   #FRK_CfgSetWalk_DeclarationUnit := FALSE;
   IF #Phase = 1 THEN
       #ConfigStageParCfg := #ParCfg;
   END_IF;
   IF #Phase = 1 THEN
       #ConfigStageStationCfg := #StationCfg;
   END_IF;
   IF "FRK_SetRuntime".Work[#RootIndex].Payload.Info.Kind = 0 THEN
       "FRK_CfgDef_DeclarationUnit"(FieldIndex := 1);
       "FRK_SetRuntime".Work[#RootIndex].RejectScope := #Status.Name;
       "FRK_SetRuntime".Work[#RootIndex].RejectKey := "FRK_ConfigScratch".Entry.WriteKey;
       IF #Phase = 0 THEN
           IF #Access.CurrentLevel < MAX(IN1 := #Access.Policy.Required[0], IN2 := "FRK_ConfigScratch".MinRead) THEN
               RETURN;
           END_IF;
           #Ok := "FRK_ConfigGet"(Scope := #Status.Name, ModelCode := "FRK_SetRuntime".Work[#RootIndex].Payload.Info.ModelCode);
           IF NOT #Ok OR "FRK_SetRuntime".Work[#RootIndex].Payload.Info.RecordCount >= 24 THEN
               RETURN;
           END_IF;
           #Slot := "FRK_SetRuntime".Work[#RootIndex].Payload.Info.RecordCount + 1;
           "FRK_SetRuntime".Work[#RootIndex].Payload.Records[#Slot].Scope := #Status.Name;
           "FRK_SetRuntime".Work[#RootIndex].Payload.Records[#Slot].WriteKey := "FRK_ConfigScratch".Entry.WriteKey;
           "FRK_SetRuntime".Work[#RootIndex].Payload.Records[#Slot].Revision := "FRK_ConfigScratch".Entry.WriteRevision;
           "FRK_SetRuntime".Work[#RootIndex].Payload.Records[#Slot].Kind := "FRK_ConfigScratch".Entry.ConfigKind;
           "FRK_SetRuntime".Work[#RootIndex].Payload.Records[#Slot].ValueType := "FRK_ConfigScratch".Entry.ValueType;
           "FRK_SetRuntime".Work[#RootIndex].Payload.Records[#Slot].ValueText := WSTRING_TO_STRING("FRK_ConfigScratch".Entry.ValueText);
           "FRK_SetRuntime".Work[#RootIndex].Payload.Info.RecordCount := #Slot;
       ELSIF #Phase = 2 THEN
           #Slot := "FRK_SetRecord"(RootIndex := #RootIndex, Scope := #Status.Name, WriteKey := "FRK_ConfigScratch".Entry.WriteKey);
           #Stored := "FRK_ConfigFind"(Scope := #Status.Name, Key := "FRK_ConfigScratch".Entry.WriteKey, ModelCode := "FRK_SetRuntime".Work[#RootIndex].Payload.Info.ModelCode);
           "FRK_ConfigStore".Rows[#Stored].Record := "FRK_SetRuntime".Work[#RootIndex].Payload.Records[#Slot];
           "FRK_ConfigStore".Rows[#Stored].SchemaVersion := "FRK_ConfigScratch".Schema;
       ELSE
           #Slot := "FRK_SetCheck"(RootIndex := #RootIndex, Scope := #Status.Name, Access := #Access, Ready := #Ready, WriteAccess := #Phase <> 3);
           IF #Slot = 0 THEN
               RETURN;
           END_IF;
           IF #Phase = 1 THEN
               #ConfigStageParCfg.Timeout := DINT_TO_TIME(LINT_TO_DINT("FRK_ConfigScratch".Value.Number));
           END_IF;
       END_IF;
   END_IF;
   IF "FRK_SetRuntime".Work[#RootIndex].Payload.Info.Kind = 0 THEN
       "FRK_CfgDef_DeclarationUnit"(FieldIndex := 2);
       "FRK_SetRuntime".Work[#RootIndex].RejectScope := #Status.Name;
       "FRK_SetRuntime".Work[#RootIndex].RejectKey := "FRK_ConfigScratch".Entry.WriteKey;
       IF #Phase = 0 THEN
           IF #Access.CurrentLevel < MAX(IN1 := #Access.Policy.Required[0], IN2 := "FRK_ConfigScratch".MinRead) THEN
               RETURN;
           END_IF;
           #Ok := "FRK_ConfigGet"(Scope := #Status.Name, ModelCode := "FRK_SetRuntime".Work[#RootIndex].Payload.Info.ModelCode);
           IF NOT #Ok OR "FRK_SetRuntime".Work[#RootIndex].Payload.Info.RecordCount >= 24 THEN
               RETURN;
           END_IF;
           #Slot := "FRK_SetRuntime".Work[#RootIndex].Payload.Info.RecordCount + 1;
           "FRK_SetRuntime".Work[#RootIndex].Payload.Records[#Slot].Scope := #Status.Name;
           "FRK_SetRuntime".Work[#RootIndex].Payload.Records[#Slot].WriteKey := "FRK_ConfigScratch".Entry.WriteKey;
           "FRK_SetRuntime".Work[#RootIndex].Payload.Records[#Slot].Revision := "FRK_ConfigScratch".Entry.WriteRevision;
           "FRK_SetRuntime".Work[#RootIndex].Payload.Records[#Slot].Kind := "FRK_ConfigScratch".Entry.ConfigKind;
           "FRK_SetRuntime".Work[#RootIndex].Payload.Records[#Slot].ValueType := "FRK_ConfigScratch".Entry.ValueType;
           "FRK_SetRuntime".Work[#RootIndex].Payload.Records[#Slot].ValueText := WSTRING_TO_STRING("FRK_ConfigScratch".Entry.ValueText);
           "FRK_SetRuntime".Work[#RootIndex].Payload.Info.RecordCount := #Slot;
       ELSIF #Phase = 2 THEN
           #Slot := "FRK_SetRecord"(RootIndex := #RootIndex, Scope := #Status.Name, WriteKey := "FRK_ConfigScratch".Entry.WriteKey);
           #Stored := "FRK_ConfigFind"(Scope := #Status.Name, Key := "FRK_ConfigScratch".Entry.WriteKey, ModelCode := "FRK_SetRuntime".Work[#RootIndex].Payload.Info.ModelCode);
           "FRK_ConfigStore".Rows[#Stored].Record := "FRK_SetRuntime".Work[#RootIndex].Payload.Records[#Slot];
           "FRK_ConfigStore".Rows[#Stored].SchemaVersion := "FRK_ConfigScratch".Schema;
       ELSE
           #Slot := "FRK_SetCheck"(RootIndex := #RootIndex, Scope := #Status.Name, Access := #Access, Ready := #Ready, WriteAccess := #Phase <> 3);
           IF #Slot = 0 THEN
               RETURN;
           END_IF;
           IF #Phase = 1 THEN
               #ConfigStageParCfg.Preset := LINT_TO_DINT("FRK_ConfigScratch".Value.Number);
           END_IF;
       END_IF;
   END_IF;
   IF "FRK_SetRuntime".Work[#RootIndex].Payload.Info.Kind = 1 THEN
       "FRK_CfgDef_DeclarationUnit"(FieldIndex := 3);
       "FRK_SetRuntime".Work[#RootIndex].RejectScope := #Status.Name;
       "FRK_SetRuntime".Work[#RootIndex].RejectKey := "FRK_ConfigScratch".Entry.WriteKey;
       IF #Phase = 0 THEN
           IF #Access.CurrentLevel < MAX(IN1 := #Access.Policy.Required[0], IN2 := "FRK_ConfigScratch".MinRead) THEN
               RETURN;
           END_IF;
           #Ok := "FRK_ConfigGet"(Scope := #Status.Name, ModelCode := "FRK_SetRuntime".Work[#RootIndex].Payload.Info.ModelCode);
           IF NOT #Ok OR "FRK_SetRuntime".Work[#RootIndex].Payload.Info.RecordCount >= 24 THEN
               RETURN;
           END_IF;
           #Slot := "FRK_SetRuntime".Work[#RootIndex].Payload.Info.RecordCount + 1;
           "FRK_SetRuntime".Work[#RootIndex].Payload.Records[#Slot].Scope := #Status.Name;
           "FRK_SetRuntime".Work[#RootIndex].Payload.Records[#Slot].WriteKey := "FRK_ConfigScratch".Entry.WriteKey;
           "FRK_SetRuntime".Work[#RootIndex].Payload.Records[#Slot].Revision := "FRK_ConfigScratch".Entry.WriteRevision;
           "FRK_SetRuntime".Work[#RootIndex].Payload.Records[#Slot].Kind := "FRK_ConfigScratch".Entry.ConfigKind;
           "FRK_SetRuntime".Work[#RootIndex].Payload.Records[#Slot].ValueType := "FRK_ConfigScratch".Entry.ValueType;
           "FRK_SetRuntime".Work[#RootIndex].Payload.Records[#Slot].ValueText := WSTRING_TO_STRING("FRK_ConfigScratch".Entry.ValueText);
           "FRK_SetRuntime".Work[#RootIndex].Payload.Info.RecordCount := #Slot;
       ELSIF #Phase = 2 THEN
           #Slot := "FRK_SetRecord"(RootIndex := #RootIndex, Scope := #Status.Name, WriteKey := "FRK_ConfigScratch".Entry.WriteKey);
           #Stored := "FRK_ConfigFind"(Scope := #Status.Name, Key := "FRK_ConfigScratch".Entry.WriteKey, ModelCode := "FRK_SetRuntime".Work[#RootIndex].Payload.Info.ModelCode);
           "FRK_ConfigStore".Rows[#Stored].Record := "FRK_SetRuntime".Work[#RootIndex].Payload.Records[#Slot];
           "FRK_ConfigStore".Rows[#Stored].SchemaVersion := "FRK_ConfigScratch".Schema;
       ELSE
           #Slot := "FRK_SetCheck"(RootIndex := #RootIndex, Scope := #Status.Name, Access := #Access, Ready := #Ready, WriteAccess := #Phase <> 3);
           IF #Slot = 0 THEN
               RETURN;
           END_IF;
           IF #Phase = 1 THEN
               #ConfigStageStationCfg.SiteLabel := "FRK_ConfigScratch".Value.Text;
           END_IF;
       END_IF;
   END_IF;
   IF "FRK_SetRuntime".Work[#RootIndex].Payload.Info.Kind = 1 THEN
       "FRK_CfgDef_DeclarationUnit"(FieldIndex := 4);
       "FRK_SetRuntime".Work[#RootIndex].RejectScope := #Status.Name;
       "FRK_SetRuntime".Work[#RootIndex].RejectKey := "FRK_ConfigScratch".Entry.WriteKey;
       IF #Phase = 0 THEN
           IF #Access.CurrentLevel < MAX(IN1 := #Access.Policy.Required[0], IN2 := "FRK_ConfigScratch".MinRead) THEN
               RETURN;
           END_IF;
           #Ok := "FRK_ConfigGet"(Scope := #Status.Name, ModelCode := "FRK_SetRuntime".Work[#RootIndex].Payload.Info.ModelCode);
           IF NOT #Ok OR "FRK_SetRuntime".Work[#RootIndex].Payload.Info.RecordCount >= 24 THEN
               RETURN;
           END_IF;
           #Slot := "FRK_SetRuntime".Work[#RootIndex].Payload.Info.RecordCount + 1;
           "FRK_SetRuntime".Work[#RootIndex].Payload.Records[#Slot].Scope := #Status.Name;
           "FRK_SetRuntime".Work[#RootIndex].Payload.Records[#Slot].WriteKey := "FRK_ConfigScratch".Entry.WriteKey;
           "FRK_SetRuntime".Work[#RootIndex].Payload.Records[#Slot].Revision := "FRK_ConfigScratch".Entry.WriteRevision;
           "FRK_SetRuntime".Work[#RootIndex].Payload.Records[#Slot].Kind := "FRK_ConfigScratch".Entry.ConfigKind;
           "FRK_SetRuntime".Work[#RootIndex].Payload.Records[#Slot].ValueType := "FRK_ConfigScratch".Entry.ValueType;
           "FRK_SetRuntime".Work[#RootIndex].Payload.Records[#Slot].ValueText := WSTRING_TO_STRING("FRK_ConfigScratch".Entry.ValueText);
           "FRK_SetRuntime".Work[#RootIndex].Payload.Info.RecordCount := #Slot;
       ELSIF #Phase = 2 THEN
           #Slot := "FRK_SetRecord"(RootIndex := #RootIndex, Scope := #Status.Name, WriteKey := "FRK_ConfigScratch".Entry.WriteKey);
           #Stored := "FRK_ConfigFind"(Scope := #Status.Name, Key := "FRK_ConfigScratch".Entry.WriteKey, ModelCode := "FRK_SetRuntime".Work[#RootIndex].Payload.Info.ModelCode);
           "FRK_ConfigStore".Rows[#Stored].Record := "FRK_SetRuntime".Work[#RootIndex].Payload.Records[#Slot];
           "FRK_ConfigStore".Rows[#Stored].SchemaVersion := "FRK_ConfigScratch".Schema;
       ELSE
           #Slot := "FRK_SetCheck"(RootIndex := #RootIndex, Scope := #Status.Name, Access := #Access, Ready := #Ready, WriteAccess := #Phase <> 3);
           IF #Slot = 0 THEN
               RETURN;
           END_IF;
           IF #Phase = 1 THEN
               #ConfigStageStationCfg.LongText := "FRK_ConfigScratch".Value.Text;
           END_IF;
       END_IF;
   END_IF;
   IF "FRK_SetRuntime".Work[#RootIndex].Payload.Info.Kind = 1 THEN
       "FRK_CfgDef_DeclarationUnit"(FieldIndex := 5);
       "FRK_SetRuntime".Work[#RootIndex].RejectScope := #Status.Name;
       "FRK_SetRuntime".Work[#RootIndex].RejectKey := "FRK_ConfigScratch".Entry.WriteKey;
       IF #Phase = 0 THEN
           IF #Access.CurrentLevel < MAX(IN1 := #Access.Policy.Required[0], IN2 := "FRK_ConfigScratch".MinRead) THEN
               RETURN;
           END_IF;
           #Ok := "FRK_ConfigGet"(Scope := #Status.Name, ModelCode := "FRK_SetRuntime".Work[#RootIndex].Payload.Info.ModelCode);
           IF NOT #Ok OR "FRK_SetRuntime".Work[#RootIndex].Payload.Info.RecordCount >= 24 THEN
               RETURN;
           END_IF;
           #Slot := "FRK_SetRuntime".Work[#RootIndex].Payload.Info.RecordCount + 1;
           "FRK_SetRuntime".Work[#RootIndex].Payload.Records[#Slot].Scope := #Status.Name;
           "FRK_SetRuntime".Work[#RootIndex].Payload.Records[#Slot].WriteKey := "FRK_ConfigScratch".Entry.WriteKey;
           "FRK_SetRuntime".Work[#RootIndex].Payload.Records[#Slot].Revision := "FRK_ConfigScratch".Entry.WriteRevision;
           "FRK_SetRuntime".Work[#RootIndex].Payload.Records[#Slot].Kind := "FRK_ConfigScratch".Entry.ConfigKind;
           "FRK_SetRuntime".Work[#RootIndex].Payload.Records[#Slot].ValueType := "FRK_ConfigScratch".Entry.ValueType;
           "FRK_SetRuntime".Work[#RootIndex].Payload.Records[#Slot].ValueText := WSTRING_TO_STRING("FRK_ConfigScratch".Entry.ValueText);
           "FRK_SetRuntime".Work[#RootIndex].Payload.Info.RecordCount := #Slot;
       ELSIF #Phase = 2 THEN
           #Slot := "FRK_SetRecord"(RootIndex := #RootIndex, Scope := #Status.Name, WriteKey := "FRK_ConfigScratch".Entry.WriteKey);
           #Stored := "FRK_ConfigFind"(Scope := #Status.Name, Key := "FRK_ConfigScratch".Entry.WriteKey, ModelCode := "FRK_SetRuntime".Work[#RootIndex].Payload.Info.ModelCode);
           "FRK_ConfigStore".Rows[#Stored].Record := "FRK_SetRuntime".Work[#RootIndex].Payload.Records[#Slot];
           "FRK_ConfigStore".Rows[#Stored].SchemaVersion := "FRK_ConfigScratch".Schema;
       ELSE
           #Slot := "FRK_SetCheck"(RootIndex := #RootIndex, Scope := #Status.Name, Access := #Access, Ready := #Ready, WriteAccess := #Phase <> 3);
           IF #Slot = 0 THEN
               RETURN;
           END_IF;
           IF #Phase = 1 THEN
               #ConfigStageStationCfg.Enabled := "FRK_ConfigScratch".Value.Flag;
           END_IF;
       END_IF;
   END_IF;
   IF #Phase = 2 AND "FRK_SetRuntime".Work[#RootIndex].Payload.Info.Kind = 0 THEN
       #ParCfg := #ConfigStageParCfg;
   END_IF;
   IF #Phase = 2 AND "FRK_SetRuntime".Work[#RootIndex].Payload.Info.Kind = 1 THEN
       #StationCfg := #ConfigStageStationCfg;
   END_IF;
   #Ok := "FRK_CfgSetWalk_DeclarationCell"(Module := #Cell, RootIndex := #RootIndex, Phase := #Phase, Access := #Access, Ready := #Ready);
   IF NOT #Ok THEN
       RETURN;
   END_IF;
   #Ok := "FRK_CfgSetWalk_SatelliteUnit"(Module := #Satellite, RootIndex := #RootIndex, Phase := #Phase, Access := #Access, Ready := #Ready);
   IF NOT #Ok THEN
       RETURN;
   END_IF;
   #FRK_CfgSetWalk_DeclarationUnit := TRUE;
END_FUNCTION

FUNCTION "FRK_CfgSetWalk_InnerUnit" : Bool   // FC146, SCL
{ S7_Optimized_Access := 'TRUE' }
VERSION : 0.1
// stored: AutoNumber true, IsIECCheckEnabled false, SetENOAutomatically false, UDAEnableTagReadback false
   VAR_INPUT
      RootIndex : Int;
      Phase : Int;
      Access : "FRK_Access";
      Ready : Bool;
   END_VAR
   VAR_IN_OUT
      Module : "FB_InnerUnit";
   END_VAR
   VAR_TEMP
      Slot : Int;
      Stored : Int;
      Ok : Bool;
   END_VAR
BEGIN

   #FRK_CfgSetWalk_InnerUnit := FALSE;
   IF #Phase = 1 THEN
       #Module.ConfigStageParCfg := #Module.ParCfg;
   END_IF;
   IF #Phase = 1 THEN
       #Module.ConfigStageStationCfg := #Module.StationCfg;
   END_IF;
   IF "FRK_SetRuntime".Work[#RootIndex].Payload.Info.Kind = 0 THEN
       "FRK_CfgDef_InnerUnit"(FieldIndex := 1);
       "FRK_SetRuntime".Work[#RootIndex].RejectScope := #Module.Status.Name;
       "FRK_SetRuntime".Work[#RootIndex].RejectKey := "FRK_ConfigScratch".Entry.WriteKey;
       IF #Phase = 0 THEN
           IF #Access.CurrentLevel < MAX(IN1 := #Access.Policy.Required[0], IN2 := "FRK_ConfigScratch".MinRead) THEN
               RETURN;
           END_IF;
           #Ok := "FRK_ConfigGet"(Scope := #Module.Status.Name, ModelCode := "FRK_SetRuntime".Work[#RootIndex].Payload.Info.ModelCode);
           IF NOT #Ok OR "FRK_SetRuntime".Work[#RootIndex].Payload.Info.RecordCount >= 24 THEN
               RETURN;
           END_IF;
           #Slot := "FRK_SetRuntime".Work[#RootIndex].Payload.Info.RecordCount + 1;
           "FRK_SetRuntime".Work[#RootIndex].Payload.Records[#Slot].Scope := #Module.Status.Name;
           "FRK_SetRuntime".Work[#RootIndex].Payload.Records[#Slot].WriteKey := "FRK_ConfigScratch".Entry.WriteKey;
           "FRK_SetRuntime".Work[#RootIndex].Payload.Records[#Slot].Revision := "FRK_ConfigScratch".Entry.WriteRevision;
           "FRK_SetRuntime".Work[#RootIndex].Payload.Records[#Slot].Kind := "FRK_ConfigScratch".Entry.ConfigKind;
           "FRK_SetRuntime".Work[#RootIndex].Payload.Records[#Slot].ValueType := "FRK_ConfigScratch".Entry.ValueType;
           "FRK_SetRuntime".Work[#RootIndex].Payload.Records[#Slot].ValueText := WSTRING_TO_STRING("FRK_ConfigScratch".Entry.ValueText);
           "FRK_SetRuntime".Work[#RootIndex].Payload.Info.RecordCount := #Slot;
       ELSIF #Phase = 2 THEN
           #Slot := "FRK_SetRecord"(RootIndex := #RootIndex, Scope := #Module.Status.Name, WriteKey := "FRK_ConfigScratch".Entry.WriteKey);
           #Stored := "FRK_ConfigFind"(Scope := #Module.Status.Name, Key := "FRK_ConfigScratch".Entry.WriteKey, ModelCode := "FRK_SetRuntime".Work[#RootIndex].Payload.Info.ModelCode);
           "FRK_ConfigStore".Rows[#Stored].Record := "FRK_SetRuntime".Work[#RootIndex].Payload.Records[#Slot];
           "FRK_ConfigStore".Rows[#Stored].SchemaVersion := "FRK_ConfigScratch".Schema;
       ELSE
           #Slot := "FRK_SetCheck"(RootIndex := #RootIndex, Scope := #Module.Status.Name, Access := #Access, Ready := #Ready, WriteAccess := #Phase <> 3);
           IF #Slot = 0 THEN
               RETURN;
           END_IF;
           IF #Phase = 1 THEN
               #Module.ConfigStageParCfg.Timeout := DINT_TO_TIME(LINT_TO_DINT("FRK_ConfigScratch".Value.Number));
           END_IF;
       END_IF;
   END_IF;
   IF "FRK_SetRuntime".Work[#RootIndex].Payload.Info.Kind = 0 THEN
       "FRK_CfgDef_InnerUnit"(FieldIndex := 2);
       "FRK_SetRuntime".Work[#RootIndex].RejectScope := #Module.Status.Name;
       "FRK_SetRuntime".Work[#RootIndex].RejectKey := "FRK_ConfigScratch".Entry.WriteKey;
       IF #Phase = 0 THEN
           IF #Access.CurrentLevel < MAX(IN1 := #Access.Policy.Required[0], IN2 := "FRK_ConfigScratch".MinRead) THEN
               RETURN;
           END_IF;
           #Ok := "FRK_ConfigGet"(Scope := #Module.Status.Name, ModelCode := "FRK_SetRuntime".Work[#RootIndex].Payload.Info.ModelCode);
           IF NOT #Ok OR "FRK_SetRuntime".Work[#RootIndex].Payload.Info.RecordCount >= 24 THEN
               RETURN;
           END_IF;
           #Slot := "FRK_SetRuntime".Work[#RootIndex].Payload.Info.RecordCount + 1;
           "FRK_SetRuntime".Work[#RootIndex].Payload.Records[#Slot].Scope := #Module.Status.Name;
           "FRK_SetRuntime".Work[#RootIndex].Payload.Records[#Slot].WriteKey := "FRK_ConfigScratch".Entry.WriteKey;
           "FRK_SetRuntime".Work[#RootIndex].Payload.Records[#Slot].Revision := "FRK_ConfigScratch".Entry.WriteRevision;
           "FRK_SetRuntime".Work[#RootIndex].Payload.Records[#Slot].Kind := "FRK_ConfigScratch".Entry.ConfigKind;
           "FRK_SetRuntime".Work[#RootIndex].Payload.Records[#Slot].ValueType := "FRK_ConfigScratch".Entry.ValueType;
           "FRK_SetRuntime".Work[#RootIndex].Payload.Records[#Slot].ValueText := WSTRING_TO_STRING("FRK_ConfigScratch".Entry.ValueText);
           "FRK_SetRuntime".Work[#RootIndex].Payload.Info.RecordCount := #Slot;
       ELSIF #Phase = 2 THEN
           #Slot := "FRK_SetRecord"(RootIndex := #RootIndex, Scope := #Module.Status.Name, WriteKey := "FRK_ConfigScratch".Entry.WriteKey);
           #Stored := "FRK_ConfigFind"(Scope := #Module.Status.Name, Key := "FRK_ConfigScratch".Entry.WriteKey, ModelCode := "FRK_SetRuntime".Work[#RootIndex].Payload.Info.ModelCode);
           "FRK_ConfigStore".Rows[#Stored].Record := "FRK_SetRuntime".Work[#RootIndex].Payload.Records[#Slot];
           "FRK_ConfigStore".Rows[#Stored].SchemaVersion := "FRK_ConfigScratch".Schema;
       ELSE
           #Slot := "FRK_SetCheck"(RootIndex := #RootIndex, Scope := #Module.Status.Name, Access := #Access, Ready := #Ready, WriteAccess := #Phase <> 3);
           IF #Slot = 0 THEN
               RETURN;
           END_IF;
           IF #Phase = 1 THEN
               #Module.ConfigStageParCfg.Preset := LINT_TO_DINT("FRK_ConfigScratch".Value.Number);
           END_IF;
       END_IF;
   END_IF;
   IF "FRK_SetRuntime".Work[#RootIndex].Payload.Info.Kind = 1 THEN
       "FRK_CfgDef_InnerUnit"(FieldIndex := 3);
       "FRK_SetRuntime".Work[#RootIndex].RejectScope := #Module.Status.Name;
       "FRK_SetRuntime".Work[#RootIndex].RejectKey := "FRK_ConfigScratch".Entry.WriteKey;
       IF #Phase = 0 THEN
           IF #Access.CurrentLevel < MAX(IN1 := #Access.Policy.Required[0], IN2 := "FRK_ConfigScratch".MinRead) THEN
               RETURN;
           END_IF;
           #Ok := "FRK_ConfigGet"(Scope := #Module.Status.Name, ModelCode := "FRK_SetRuntime".Work[#RootIndex].Payload.Info.ModelCode);
           IF NOT #Ok OR "FRK_SetRuntime".Work[#RootIndex].Payload.Info.RecordCount >= 24 THEN
               RETURN;
           END_IF;
           #Slot := "FRK_SetRuntime".Work[#RootIndex].Payload.Info.RecordCount + 1;
           "FRK_SetRuntime".Work[#RootIndex].Payload.Records[#Slot].Scope := #Module.Status.Name;
           "FRK_SetRuntime".Work[#RootIndex].Payload.Records[#Slot].WriteKey := "FRK_ConfigScratch".Entry.WriteKey;
           "FRK_SetRuntime".Work[#RootIndex].Payload.Records[#Slot].Revision := "FRK_ConfigScratch".Entry.WriteRevision;
           "FRK_SetRuntime".Work[#RootIndex].Payload.Records[#Slot].Kind := "FRK_ConfigScratch".Entry.ConfigKind;
           "FRK_SetRuntime".Work[#RootIndex].Payload.Records[#Slot].ValueType := "FRK_ConfigScratch".Entry.ValueType;
           "FRK_SetRuntime".Work[#RootIndex].Payload.Records[#Slot].ValueText := WSTRING_TO_STRING("FRK_ConfigScratch".Entry.ValueText);
           "FRK_SetRuntime".Work[#RootIndex].Payload.Info.RecordCount := #Slot;
       ELSIF #Phase = 2 THEN
           #Slot := "FRK_SetRecord"(RootIndex := #RootIndex, Scope := #Module.Status.Name, WriteKey := "FRK_ConfigScratch".Entry.WriteKey);
           #Stored := "FRK_ConfigFind"(Scope := #Module.Status.Name, Key := "FRK_ConfigScratch".Entry.WriteKey, ModelCode := "FRK_SetRuntime".Work[#RootIndex].Payload.Info.ModelCode);
           "FRK_ConfigStore".Rows[#Stored].Record := "FRK_SetRuntime".Work[#RootIndex].Payload.Records[#Slot];
           "FRK_ConfigStore".Rows[#Stored].SchemaVersion := "FRK_ConfigScratch".Schema;
       ELSE
           #Slot := "FRK_SetCheck"(RootIndex := #RootIndex, Scope := #Module.Status.Name, Access := #Access, Ready := #Ready, WriteAccess := #Phase <> 3);
           IF #Slot = 0 THEN
               RETURN;
           END_IF;
           IF #Phase = 1 THEN
               #Module.ConfigStageStationCfg.SiteLabel := "FRK_ConfigScratch".Value.Text;
           END_IF;
       END_IF;
   END_IF;
   IF "FRK_SetRuntime".Work[#RootIndex].Payload.Info.Kind = 1 THEN
       "FRK_CfgDef_InnerUnit"(FieldIndex := 4);
       "FRK_SetRuntime".Work[#RootIndex].RejectScope := #Module.Status.Name;
       "FRK_SetRuntime".Work[#RootIndex].RejectKey := "FRK_ConfigScratch".Entry.WriteKey;
       IF #Phase = 0 THEN
           IF #Access.CurrentLevel < MAX(IN1 := #Access.Policy.Required[0], IN2 := "FRK_ConfigScratch".MinRead) THEN
               RETURN;
           END_IF;
           #Ok := "FRK_ConfigGet"(Scope := #Module.Status.Name, ModelCode := "FRK_SetRuntime".Work[#RootIndex].Payload.Info.ModelCode);
           IF NOT #Ok OR "FRK_SetRuntime".Work[#RootIndex].Payload.Info.RecordCount >= 24 THEN
               RETURN;
           END_IF;
           #Slot := "FRK_SetRuntime".Work[#RootIndex].Payload.Info.RecordCount + 1;
           "FRK_SetRuntime".Work[#RootIndex].Payload.Records[#Slot].Scope := #Module.Status.Name;
           "FRK_SetRuntime".Work[#RootIndex].Payload.Records[#Slot].WriteKey := "FRK_ConfigScratch".Entry.WriteKey;
           "FRK_SetRuntime".Work[#RootIndex].Payload.Records[#Slot].Revision := "FRK_ConfigScratch".Entry.WriteRevision;
           "FRK_SetRuntime".Work[#RootIndex].Payload.Records[#Slot].Kind := "FRK_ConfigScratch".Entry.ConfigKind;
           "FRK_SetRuntime".Work[#RootIndex].Payload.Records[#Slot].ValueType := "FRK_ConfigScratch".Entry.ValueType;
           "FRK_SetRuntime".Work[#RootIndex].Payload.Records[#Slot].ValueText := WSTRING_TO_STRING("FRK_ConfigScratch".Entry.ValueText);
           "FRK_SetRuntime".Work[#RootIndex].Payload.Info.RecordCount := #Slot;
       ELSIF #Phase = 2 THEN
           #Slot := "FRK_SetRecord"(RootIndex := #RootIndex, Scope := #Module.Status.Name, WriteKey := "FRK_ConfigScratch".Entry.WriteKey);
           #Stored := "FRK_ConfigFind"(Scope := #Module.Status.Name, Key := "FRK_ConfigScratch".Entry.WriteKey, ModelCode := "FRK_SetRuntime".Work[#RootIndex].Payload.Info.ModelCode);
           "FRK_ConfigStore".Rows[#Stored].Record := "FRK_SetRuntime".Work[#RootIndex].Payload.Records[#Slot];
           "FRK_ConfigStore".Rows[#Stored].SchemaVersion := "FRK_ConfigScratch".Schema;
       ELSE
           #Slot := "FRK_SetCheck"(RootIndex := #RootIndex, Scope := #Module.Status.Name, Access := #Access, Ready := #Ready, WriteAccess := #Phase <> 3);
           IF #Slot = 0 THEN
               RETURN;
           END_IF;
           IF #Phase = 1 THEN
               #Module.ConfigStageStationCfg.LongText := "FRK_ConfigScratch".Value.Text;
           END_IF;
       END_IF;
   END_IF;
   IF "FRK_SetRuntime".Work[#RootIndex].Payload.Info.Kind = 1 THEN
       "FRK_CfgDef_InnerUnit"(FieldIndex := 5);
       "FRK_SetRuntime".Work[#RootIndex].RejectScope := #Module.Status.Name;
       "FRK_SetRuntime".Work[#RootIndex].RejectKey := "FRK_ConfigScratch".Entry.WriteKey;
       IF #Phase = 0 THEN
           IF #Access.CurrentLevel < MAX(IN1 := #Access.Policy.Required[0], IN2 := "FRK_ConfigScratch".MinRead) THEN
               RETURN;
           END_IF;
           #Ok := "FRK_ConfigGet"(Scope := #Module.Status.Name, ModelCode := "FRK_SetRuntime".Work[#RootIndex].Payload.Info.ModelCode);
           IF NOT #Ok OR "FRK_SetRuntime".Work[#RootIndex].Payload.Info.RecordCount >= 24 THEN
               RETURN;
           END_IF;
           #Slot := "FRK_SetRuntime".Work[#RootIndex].Payload.Info.RecordCount + 1;
           "FRK_SetRuntime".Work[#RootIndex].Payload.Records[#Slot].Scope := #Module.Status.Name;
           "FRK_SetRuntime".Work[#RootIndex].Payload.Records[#Slot].WriteKey := "FRK_ConfigScratch".Entry.WriteKey;
           "FRK_SetRuntime".Work[#RootIndex].Payload.Records[#Slot].Revision := "FRK_ConfigScratch".Entry.WriteRevision;
           "FRK_SetRuntime".Work[#RootIndex].Payload.Records[#Slot].Kind := "FRK_ConfigScratch".Entry.ConfigKind;
           "FRK_SetRuntime".Work[#RootIndex].Payload.Records[#Slot].ValueType := "FRK_ConfigScratch".Entry.ValueType;
           "FRK_SetRuntime".Work[#RootIndex].Payload.Records[#Slot].ValueText := WSTRING_TO_STRING("FRK_ConfigScratch".Entry.ValueText);
           "FRK_SetRuntime".Work[#RootIndex].Payload.Info.RecordCount := #Slot;
       ELSIF #Phase = 2 THEN
           #Slot := "FRK_SetRecord"(RootIndex := #RootIndex, Scope := #Module.Status.Name, WriteKey := "FRK_ConfigScratch".Entry.WriteKey);
           #Stored := "FRK_ConfigFind"(Scope := #Module.Status.Name, Key := "FRK_ConfigScratch".Entry.WriteKey, ModelCode := "FRK_SetRuntime".Work[#RootIndex].Payload.Info.ModelCode);
           "FRK_ConfigStore".Rows[#Stored].Record := "FRK_SetRuntime".Work[#RootIndex].Payload.Records[#Slot];
           "FRK_ConfigStore".Rows[#Stored].SchemaVersion := "FRK_ConfigScratch".Schema;
       ELSE
           #Slot := "FRK_SetCheck"(RootIndex := #RootIndex, Scope := #Module.Status.Name, Access := #Access, Ready := #Ready, WriteAccess := #Phase <> 3);
           IF #Slot = 0 THEN
               RETURN;
           END_IF;
           IF #Phase = 1 THEN
               #Module.ConfigStageStationCfg.Enabled := "FRK_ConfigScratch".Value.Flag;
           END_IF;
       END_IF;
   END_IF;
   IF #Phase = 2 AND "FRK_SetRuntime".Work[#RootIndex].Payload.Info.Kind = 0 THEN
       #Module.ParCfg := #Module.ConfigStageParCfg;
   END_IF;
   IF #Phase = 2 AND "FRK_SetRuntime".Work[#RootIndex].Payload.Info.Kind = 1 THEN
       #Module.StationCfg := #Module.ConfigStageStationCfg;
   END_IF;
   #Ok := "FRK_CfgSetWalk_DeclarationCell"(Module := #Module.Cell, RootIndex := #RootIndex, Phase := #Phase, Access := #Access, Ready := #Ready);
   IF NOT #Ok THEN
       RETURN;
   END_IF;
   #FRK_CfgSetWalk_InnerUnit := TRUE;
END_FUNCTION

FUNCTION "FRK_CfgSetWalk_SatelliteUnit" : Bool   // FC154, SCL
{ S7_Optimized_Access := 'TRUE' }
VERSION : 0.1
// stored: AutoNumber true, IsIECCheckEnabled false, SetENOAutomatically false, UDAEnableTagReadback false
   VAR_INPUT
      RootIndex : Int;
      Phase : Int;
      Access : "FRK_Access";
      Ready : Bool;
   END_VAR
   VAR_IN_OUT
      Module : "FB_SatelliteUnit";
   END_VAR
   VAR_TEMP
      Slot : Int;
      Stored : Int;
      Ok : Bool;
   END_VAR
BEGIN

   #FRK_CfgSetWalk_SatelliteUnit := FALSE;
   IF #Phase = 1 THEN
       #Module.ConfigStageParCfg := #Module.ParCfg;
   END_IF;
   IF #Phase = 1 THEN
       #Module.ConfigStageStationCfg := #Module.StationCfg;
   END_IF;
   IF "FRK_SetRuntime".Work[#RootIndex].Payload.Info.Kind = 0 THEN
       "FRK_CfgDef_SatelliteUnit"(FieldIndex := 1);
       "FRK_SetRuntime".Work[#RootIndex].RejectScope := #Module.Status.Name;
       "FRK_SetRuntime".Work[#RootIndex].RejectKey := "FRK_ConfigScratch".Entry.WriteKey;
       IF #Phase = 0 THEN
           IF #Access.CurrentLevel < MAX(IN1 := #Access.Policy.Required[0], IN2 := "FRK_ConfigScratch".MinRead) THEN
               RETURN;
           END_IF;
           #Ok := "FRK_ConfigGet"(Scope := #Module.Status.Name, ModelCode := "FRK_SetRuntime".Work[#RootIndex].Payload.Info.ModelCode);
           IF NOT #Ok OR "FRK_SetRuntime".Work[#RootIndex].Payload.Info.RecordCount >= 24 THEN
               RETURN;
           END_IF;
           #Slot := "FRK_SetRuntime".Work[#RootIndex].Payload.Info.RecordCount + 1;
           "FRK_SetRuntime".Work[#RootIndex].Payload.Records[#Slot].Scope := #Module.Status.Name;
           "FRK_SetRuntime".Work[#RootIndex].Payload.Records[#Slot].WriteKey := "FRK_ConfigScratch".Entry.WriteKey;
           "FRK_SetRuntime".Work[#RootIndex].Payload.Records[#Slot].Revision := "FRK_ConfigScratch".Entry.WriteRevision;
           "FRK_SetRuntime".Work[#RootIndex].Payload.Records[#Slot].Kind := "FRK_ConfigScratch".Entry.ConfigKind;
           "FRK_SetRuntime".Work[#RootIndex].Payload.Records[#Slot].ValueType := "FRK_ConfigScratch".Entry.ValueType;
           "FRK_SetRuntime".Work[#RootIndex].Payload.Records[#Slot].ValueText := WSTRING_TO_STRING("FRK_ConfigScratch".Entry.ValueText);
           "FRK_SetRuntime".Work[#RootIndex].Payload.Info.RecordCount := #Slot;
       ELSIF #Phase = 2 THEN
           #Slot := "FRK_SetRecord"(RootIndex := #RootIndex, Scope := #Module.Status.Name, WriteKey := "FRK_ConfigScratch".Entry.WriteKey);
           #Stored := "FRK_ConfigFind"(Scope := #Module.Status.Name, Key := "FRK_ConfigScratch".Entry.WriteKey, ModelCode := "FRK_SetRuntime".Work[#RootIndex].Payload.Info.ModelCode);
           "FRK_ConfigStore".Rows[#Stored].Record := "FRK_SetRuntime".Work[#RootIndex].Payload.Records[#Slot];
           "FRK_ConfigStore".Rows[#Stored].SchemaVersion := "FRK_ConfigScratch".Schema;
       ELSE
           #Slot := "FRK_SetCheck"(RootIndex := #RootIndex, Scope := #Module.Status.Name, Access := #Access, Ready := #Ready, WriteAccess := #Phase <> 3);
           IF #Slot = 0 THEN
               RETURN;
           END_IF;
           IF #Phase = 1 THEN
               #Module.ConfigStageParCfg.Timeout := DINT_TO_TIME(LINT_TO_DINT("FRK_ConfigScratch".Value.Number));
           END_IF;
       END_IF;
   END_IF;
   IF "FRK_SetRuntime".Work[#RootIndex].Payload.Info.Kind = 0 THEN
       "FRK_CfgDef_SatelliteUnit"(FieldIndex := 2);
       "FRK_SetRuntime".Work[#RootIndex].RejectScope := #Module.Status.Name;
       "FRK_SetRuntime".Work[#RootIndex].RejectKey := "FRK_ConfigScratch".Entry.WriteKey;
       IF #Phase = 0 THEN
           IF #Access.CurrentLevel < MAX(IN1 := #Access.Policy.Required[0], IN2 := "FRK_ConfigScratch".MinRead) THEN
               RETURN;
           END_IF;
           #Ok := "FRK_ConfigGet"(Scope := #Module.Status.Name, ModelCode := "FRK_SetRuntime".Work[#RootIndex].Payload.Info.ModelCode);
           IF NOT #Ok OR "FRK_SetRuntime".Work[#RootIndex].Payload.Info.RecordCount >= 24 THEN
               RETURN;
           END_IF;
           #Slot := "FRK_SetRuntime".Work[#RootIndex].Payload.Info.RecordCount + 1;
           "FRK_SetRuntime".Work[#RootIndex].Payload.Records[#Slot].Scope := #Module.Status.Name;
           "FRK_SetRuntime".Work[#RootIndex].Payload.Records[#Slot].WriteKey := "FRK_ConfigScratch".Entry.WriteKey;
           "FRK_SetRuntime".Work[#RootIndex].Payload.Records[#Slot].Revision := "FRK_ConfigScratch".Entry.WriteRevision;
           "FRK_SetRuntime".Work[#RootIndex].Payload.Records[#Slot].Kind := "FRK_ConfigScratch".Entry.ConfigKind;
           "FRK_SetRuntime".Work[#RootIndex].Payload.Records[#Slot].ValueType := "FRK_ConfigScratch".Entry.ValueType;
           "FRK_SetRuntime".Work[#RootIndex].Payload.Records[#Slot].ValueText := WSTRING_TO_STRING("FRK_ConfigScratch".Entry.ValueText);
           "FRK_SetRuntime".Work[#RootIndex].Payload.Info.RecordCount := #Slot;
       ELSIF #Phase = 2 THEN
           #Slot := "FRK_SetRecord"(RootIndex := #RootIndex, Scope := #Module.Status.Name, WriteKey := "FRK_ConfigScratch".Entry.WriteKey);
           #Stored := "FRK_ConfigFind"(Scope := #Module.Status.Name, Key := "FRK_ConfigScratch".Entry.WriteKey, ModelCode := "FRK_SetRuntime".Work[#RootIndex].Payload.Info.ModelCode);
           "FRK_ConfigStore".Rows[#Stored].Record := "FRK_SetRuntime".Work[#RootIndex].Payload.Records[#Slot];
           "FRK_ConfigStore".Rows[#Stored].SchemaVersion := "FRK_ConfigScratch".Schema;
       ELSE
           #Slot := "FRK_SetCheck"(RootIndex := #RootIndex, Scope := #Module.Status.Name, Access := #Access, Ready := #Ready, WriteAccess := #Phase <> 3);
           IF #Slot = 0 THEN
               RETURN;
           END_IF;
           IF #Phase = 1 THEN
               #Module.ConfigStageParCfg.Preset := LINT_TO_DINT("FRK_ConfigScratch".Value.Number);
           END_IF;
       END_IF;
   END_IF;
   IF "FRK_SetRuntime".Work[#RootIndex].Payload.Info.Kind = 1 THEN
       "FRK_CfgDef_SatelliteUnit"(FieldIndex := 3);
       "FRK_SetRuntime".Work[#RootIndex].RejectScope := #Module.Status.Name;
       "FRK_SetRuntime".Work[#RootIndex].RejectKey := "FRK_ConfigScratch".Entry.WriteKey;
       IF #Phase = 0 THEN
           IF #Access.CurrentLevel < MAX(IN1 := #Access.Policy.Required[0], IN2 := "FRK_ConfigScratch".MinRead) THEN
               RETURN;
           END_IF;
           #Ok := "FRK_ConfigGet"(Scope := #Module.Status.Name, ModelCode := "FRK_SetRuntime".Work[#RootIndex].Payload.Info.ModelCode);
           IF NOT #Ok OR "FRK_SetRuntime".Work[#RootIndex].Payload.Info.RecordCount >= 24 THEN
               RETURN;
           END_IF;
           #Slot := "FRK_SetRuntime".Work[#RootIndex].Payload.Info.RecordCount + 1;
           "FRK_SetRuntime".Work[#RootIndex].Payload.Records[#Slot].Scope := #Module.Status.Name;
           "FRK_SetRuntime".Work[#RootIndex].Payload.Records[#Slot].WriteKey := "FRK_ConfigScratch".Entry.WriteKey;
           "FRK_SetRuntime".Work[#RootIndex].Payload.Records[#Slot].Revision := "FRK_ConfigScratch".Entry.WriteRevision;
           "FRK_SetRuntime".Work[#RootIndex].Payload.Records[#Slot].Kind := "FRK_ConfigScratch".Entry.ConfigKind;
           "FRK_SetRuntime".Work[#RootIndex].Payload.Records[#Slot].ValueType := "FRK_ConfigScratch".Entry.ValueType;
           "FRK_SetRuntime".Work[#RootIndex].Payload.Records[#Slot].ValueText := WSTRING_TO_STRING("FRK_ConfigScratch".Entry.ValueText);
           "FRK_SetRuntime".Work[#RootIndex].Payload.Info.RecordCount := #Slot;
       ELSIF #Phase = 2 THEN
           #Slot := "FRK_SetRecord"(RootIndex := #RootIndex, Scope := #Module.Status.Name, WriteKey := "FRK_ConfigScratch".Entry.WriteKey);
           #Stored := "FRK_ConfigFind"(Scope := #Module.Status.Name, Key := "FRK_ConfigScratch".Entry.WriteKey, ModelCode := "FRK_SetRuntime".Work[#RootIndex].Payload.Info.ModelCode);
           "FRK_ConfigStore".Rows[#Stored].Record := "FRK_SetRuntime".Work[#RootIndex].Payload.Records[#Slot];
           "FRK_ConfigStore".Rows[#Stored].SchemaVersion := "FRK_ConfigScratch".Schema;
       ELSE
           #Slot := "FRK_SetCheck"(RootIndex := #RootIndex, Scope := #Module.Status.Name, Access := #Access, Ready := #Ready, WriteAccess := #Phase <> 3);
           IF #Slot = 0 THEN
               RETURN;
           END_IF;
           IF #Phase = 1 THEN
               #Module.ConfigStageStationCfg.SiteLabel := "FRK_ConfigScratch".Value.Text;
           END_IF;
       END_IF;
   END_IF;
   IF "FRK_SetRuntime".Work[#RootIndex].Payload.Info.Kind = 1 THEN
       "FRK_CfgDef_SatelliteUnit"(FieldIndex := 4);
       "FRK_SetRuntime".Work[#RootIndex].RejectScope := #Module.Status.Name;
       "FRK_SetRuntime".Work[#RootIndex].RejectKey := "FRK_ConfigScratch".Entry.WriteKey;
       IF #Phase = 0 THEN
           IF #Access.CurrentLevel < MAX(IN1 := #Access.Policy.Required[0], IN2 := "FRK_ConfigScratch".MinRead) THEN
               RETURN;
           END_IF;
           #Ok := "FRK_ConfigGet"(Scope := #Module.Status.Name, ModelCode := "FRK_SetRuntime".Work[#RootIndex].Payload.Info.ModelCode);
           IF NOT #Ok OR "FRK_SetRuntime".Work[#RootIndex].Payload.Info.RecordCount >= 24 THEN
               RETURN;
           END_IF;
           #Slot := "FRK_SetRuntime".Work[#RootIndex].Payload.Info.RecordCount + 1;
           "FRK_SetRuntime".Work[#RootIndex].Payload.Records[#Slot].Scope := #Module.Status.Name;
           "FRK_SetRuntime".Work[#RootIndex].Payload.Records[#Slot].WriteKey := "FRK_ConfigScratch".Entry.WriteKey;
           "FRK_SetRuntime".Work[#RootIndex].Payload.Records[#Slot].Revision := "FRK_ConfigScratch".Entry.WriteRevision;
           "FRK_SetRuntime".Work[#RootIndex].Payload.Records[#Slot].Kind := "FRK_ConfigScratch".Entry.ConfigKind;
           "FRK_SetRuntime".Work[#RootIndex].Payload.Records[#Slot].ValueType := "FRK_ConfigScratch".Entry.ValueType;
           "FRK_SetRuntime".Work[#RootIndex].Payload.Records[#Slot].ValueText := WSTRING_TO_STRING("FRK_ConfigScratch".Entry.ValueText);
           "FRK_SetRuntime".Work[#RootIndex].Payload.Info.RecordCount := #Slot;
       ELSIF #Phase = 2 THEN
           #Slot := "FRK_SetRecord"(RootIndex := #RootIndex, Scope := #Module.Status.Name, WriteKey := "FRK_ConfigScratch".Entry.WriteKey);
           #Stored := "FRK_ConfigFind"(Scope := #Module.Status.Name, Key := "FRK_ConfigScratch".Entry.WriteKey, ModelCode := "FRK_SetRuntime".Work[#RootIndex].Payload.Info.ModelCode);
           "FRK_ConfigStore".Rows[#Stored].Record := "FRK_SetRuntime".Work[#RootIndex].Payload.Records[#Slot];
           "FRK_ConfigStore".Rows[#Stored].SchemaVersion := "FRK_ConfigScratch".Schema;
       ELSE
           #Slot := "FRK_SetCheck"(RootIndex := #RootIndex, Scope := #Module.Status.Name, Access := #Access, Ready := #Ready, WriteAccess := #Phase <> 3);
           IF #Slot = 0 THEN
               RETURN;
           END_IF;
           IF #Phase = 1 THEN
               #Module.ConfigStageStationCfg.LongText := "FRK_ConfigScratch".Value.Text;
           END_IF;
       END_IF;
   END_IF;
   IF "FRK_SetRuntime".Work[#RootIndex].Payload.Info.Kind = 1 THEN
       "FRK_CfgDef_SatelliteUnit"(FieldIndex := 5);
       "FRK_SetRuntime".Work[#RootIndex].RejectScope := #Module.Status.Name;
       "FRK_SetRuntime".Work[#RootIndex].RejectKey := "FRK_ConfigScratch".Entry.WriteKey;
       IF #Phase = 0 THEN
           IF #Access.CurrentLevel < MAX(IN1 := #Access.Policy.Required[0], IN2 := "FRK_ConfigScratch".MinRead) THEN
               RETURN;
           END_IF;
           #Ok := "FRK_ConfigGet"(Scope := #Module.Status.Name, ModelCode := "FRK_SetRuntime".Work[#RootIndex].Payload.Info.ModelCode);
           IF NOT #Ok OR "FRK_SetRuntime".Work[#RootIndex].Payload.Info.RecordCount >= 24 THEN
               RETURN;
           END_IF;
           #Slot := "FRK_SetRuntime".Work[#RootIndex].Payload.Info.RecordCount + 1;
           "FRK_SetRuntime".Work[#RootIndex].Payload.Records[#Slot].Scope := #Module.Status.Name;
           "FRK_SetRuntime".Work[#RootIndex].Payload.Records[#Slot].WriteKey := "FRK_ConfigScratch".Entry.WriteKey;
           "FRK_SetRuntime".Work[#RootIndex].Payload.Records[#Slot].Revision := "FRK_ConfigScratch".Entry.WriteRevision;
           "FRK_SetRuntime".Work[#RootIndex].Payload.Records[#Slot].Kind := "FRK_ConfigScratch".Entry.ConfigKind;
           "FRK_SetRuntime".Work[#RootIndex].Payload.Records[#Slot].ValueType := "FRK_ConfigScratch".Entry.ValueType;
           "FRK_SetRuntime".Work[#RootIndex].Payload.Records[#Slot].ValueText := WSTRING_TO_STRING("FRK_ConfigScratch".Entry.ValueText);
           "FRK_SetRuntime".Work[#RootIndex].Payload.Info.RecordCount := #Slot;
       ELSIF #Phase = 2 THEN
           #Slot := "FRK_SetRecord"(RootIndex := #RootIndex, Scope := #Module.Status.Name, WriteKey := "FRK_ConfigScratch".Entry.WriteKey);
           #Stored := "FRK_ConfigFind"(Scope := #Module.Status.Name, Key := "FRK_ConfigScratch".Entry.WriteKey, ModelCode := "FRK_SetRuntime".Work[#RootIndex].Payload.Info.ModelCode);
           "FRK_ConfigStore".Rows[#Stored].Record := "FRK_SetRuntime".Work[#RootIndex].Payload.Records[#Slot];
           "FRK_ConfigStore".Rows[#Stored].SchemaVersion := "FRK_ConfigScratch".Schema;
       ELSE
           #Slot := "FRK_SetCheck"(RootIndex := #RootIndex, Scope := #Module.Status.Name, Access := #Access, Ready := #Ready, WriteAccess := #Phase <> 3);
           IF #Slot = 0 THEN
               RETURN;
           END_IF;
           IF #Phase = 1 THEN
               #Module.ConfigStageStationCfg.Enabled := "FRK_ConfigScratch".Value.Flag;
           END_IF;
       END_IF;
   END_IF;
   IF #Phase = 2 AND "FRK_SetRuntime".Work[#RootIndex].Payload.Info.Kind = 0 THEN
       #Module.ParCfg := #Module.ConfigStageParCfg;
   END_IF;
   IF #Phase = 2 AND "FRK_SetRuntime".Work[#RootIndex].Payload.Info.Kind = 1 THEN
       #Module.StationCfg := #Module.ConfigStageStationCfg;
   END_IF;
   #Ok := "FRK_CfgSetWalk_DeclarationCell"(Module := #Module.Cell, RootIndex := #RootIndex, Phase := #Phase, Access := #Access, Ready := #Ready);
   IF NOT #Ok THEN
       RETURN;
   END_IF;
   #Ok := "FRK_CfgSetWalk_InnerUnit"(Module := #Module.Inner, RootIndex := #RootIndex, Phase := #Phase, Access := #Access, Ready := #Ready);
   IF NOT #Ok THEN
       RETURN;
   END_IF;
   #FRK_CfgSetWalk_SatelliteUnit := TRUE;
END_FUNCTION

FUNCTION "FRK_CfgWrite_DeclarationCell" : Bool   // FC135, SCL
{ S7_Optimized_Access := 'TRUE' }
VERSION : 0.1
// stored: AutoNumber true, IsIECCheckEnabled false, SetENOAutomatically false, UDAEnableTagReadback false
   VAR_INPUT
      Request : "ST_HmiRequest";
      Access : "FRK_Access";
      RootIndex : Int;
      RootReady : Bool;
   END_VAR
   VAR_IN_OUT
      Module : "FB_DeclarationCell";
      Matched : Bool;
   END_VAR
   VAR_TEMP
      Ok : Bool;
      Level : DInt;
      Code : String[64];
      Inactive : Bool;
   END_VAR
BEGIN

   #FRK_CfgWrite_DeclarationCell := FALSE;
   IF #Request.TargetPath = STRING_TO_WSTRING(#Module.Status.Name) OR (#Request.TargetPath = WSTRING#'' AND #Module.Core.ParentIndex = 0) THEN
       "FRK_CfgDef_DeclarationCell"(FieldIndex := 1);
       IF #Request.NameValue = "FRK_ConfigScratch".Entry.WriteKey THEN
           #Matched := TRUE;
           IF DINT_TO_UDINT(#Request.IntValue) <> "FRK_ConfigScratch".Entry.WriteRevision THEN
               RETURN;
           END_IF;
           #Level := MAX(IN1 := #Access.Policy.Required[1], IN2 := "FRK_ConfigScratch".MinWrite);
           IF #Access.CurrentLevel < #Level THEN
               RETURN;
           END_IF;
           IF #Request.DurationMs <> 0 THEN
               RETURN;
           END_IF;
           #Code := "FRK_ConfigModelCode"(RootIndex := #RootIndex, ModelIndex := #Request.DurationMs);
           #Inactive := #Code <> "FRK_ConfigStore".ActiveModels[#RootIndex];
           IF "FRK_ConfigScratch".Entry.RequiresReady AND NOT #Inactive AND NOT #RootReady THEN
               RETURN;
           END_IF;
           #Ok := "FRK_ConfigDecode"(Text := #Request.TextValue, Storage := "FRK_ConfigScratch".Storage, Minimum := "FRK_ConfigScratch".Minimum, Maximum := "FRK_ConfigScratch".Maximum, MaxLength := "FRK_ConfigScratch".MaxLength, Value := "FRK_ConfigScratch".Value);
           IF NOT #Ok THEN
               RETURN;
           END_IF;
           #Ok := "FRK_ConfigPut"(Scope := #Module.Status.Name, ModelCode := #Code, Text := #Request.TextValue, RootIndex := #RootIndex);
           IF NOT #Ok THEN
               RETURN;
           END_IF;
           IF NOT #Inactive THEN
               #Module.ParCfg.Timeout := DINT_TO_TIME(LINT_TO_DINT("FRK_ConfigScratch".Value.Number));
           END_IF;
           #FRK_CfgWrite_DeclarationCell := TRUE;
           RETURN;
       END_IF;
       "FRK_CfgDef_DeclarationCell"(FieldIndex := 2);
       IF #Request.NameValue = "FRK_ConfigScratch".Entry.WriteKey THEN
           #Matched := TRUE;
           IF DINT_TO_UDINT(#Request.IntValue) <> "FRK_ConfigScratch".Entry.WriteRevision THEN
               RETURN;
           END_IF;
           #Level := MAX(IN1 := #Access.Policy.Required[1], IN2 := "FRK_ConfigScratch".MinWrite);
           IF #Access.CurrentLevel < #Level THEN
               RETURN;
           END_IF;
           IF #Request.DurationMs <> 0 THEN
               RETURN;
           END_IF;
           #Code := "FRK_ConfigModelCode"(RootIndex := #RootIndex, ModelIndex := #Request.DurationMs);
           #Inactive := #Code <> "FRK_ConfigStore".ActiveModels[#RootIndex];
           IF "FRK_ConfigScratch".Entry.RequiresReady AND NOT #Inactive AND NOT #RootReady THEN
               RETURN;
           END_IF;
           #Ok := "FRK_ConfigDecode"(Text := #Request.TextValue, Storage := "FRK_ConfigScratch".Storage, Minimum := "FRK_ConfigScratch".Minimum, Maximum := "FRK_ConfigScratch".Maximum, MaxLength := "FRK_ConfigScratch".MaxLength, Value := "FRK_ConfigScratch".Value);
           IF NOT #Ok THEN
               RETURN;
           END_IF;
           #Ok := "FRK_ConfigPut"(Scope := #Module.Status.Name, ModelCode := #Code, Text := #Request.TextValue, RootIndex := #RootIndex);
           IF NOT #Ok THEN
               RETURN;
           END_IF;
           IF NOT #Inactive THEN
               #Module.ParCfg.Preset := LINT_TO_DINT("FRK_ConfigScratch".Value.Number);
           END_IF;
           #FRK_CfgWrite_DeclarationCell := TRUE;
           RETURN;
       END_IF;
   END_IF;
   #Ok := "FRK_CfgWrite_DeclarationCylinder"(Module := #Module.Clamp, Access := #Access, Request := #Request, RootIndex := #RootIndex, RootReady := #RootReady, Matched := #Matched);
   IF #Matched THEN
       #FRK_CfgWrite_DeclarationCell := #Ok;
       RETURN;
   END_IF;
   #Ok := "FRK_CfgWrite_DeclarationCylinder"(Module := #Module.Gate, Access := #Access, Request := #Request, RootIndex := #RootIndex, RootReady := #RootReady, Matched := #Matched);
   IF #Matched THEN
       #FRK_CfgWrite_DeclarationCell := #Ok;
       RETURN;
   END_IF;
END_FUNCTION

FUNCTION "FRK_CfgWrite_DeclarationCylinder" : Bool   // FC127, SCL
{ S7_Optimized_Access := 'TRUE' }
VERSION : 0.1
// stored: AutoNumber true, IsIECCheckEnabled false, SetENOAutomatically false, UDAEnableTagReadback false
   VAR_INPUT
      Request : "ST_HmiRequest";
      Access : "FRK_Access";
      RootIndex : Int;
      RootReady : Bool;
   END_VAR
   VAR_IN_OUT
      Module : "FB_DeclarationCylinder";
      Matched : Bool;
   END_VAR
   VAR_TEMP
      Ok : Bool;
      Level : DInt;
      Code : String[64];
      Inactive : Bool;
   END_VAR
BEGIN

   #FRK_CfgWrite_DeclarationCylinder := FALSE;
   IF #Request.TargetPath = STRING_TO_WSTRING(#Module.Status.Name) OR (#Request.TargetPath = WSTRING#'' AND #Module.Core.ParentIndex = 0) THEN
       "FRK_CfgDef_DeclarationCylinder"(FieldIndex := 1);
       IF #Request.NameValue = "FRK_ConfigScratch".Entry.WriteKey THEN
           #Matched := TRUE;
           IF DINT_TO_UDINT(#Request.IntValue) <> "FRK_ConfigScratch".Entry.WriteRevision THEN
               RETURN;
           END_IF;
           #Level := MAX(IN1 := #Access.Policy.Required[1], IN2 := "FRK_ConfigScratch".MinWrite);
           IF #Access.CurrentLevel < #Level THEN
               RETURN;
           END_IF;
           IF #Request.DurationMs <> 0 THEN
               RETURN;
           END_IF;
           #Code := "FRK_ConfigModelCode"(RootIndex := #RootIndex, ModelIndex := #Request.DurationMs);
           #Inactive := #Code <> "FRK_ConfigStore".ActiveModels[#RootIndex];
           IF "FRK_ConfigScratch".Entry.RequiresReady AND NOT #Inactive AND NOT #RootReady THEN
               RETURN;
           END_IF;
           #Ok := "FRK_ConfigDecode"(Text := #Request.TextValue, Storage := "FRK_ConfigScratch".Storage, Minimum := "FRK_ConfigScratch".Minimum, Maximum := "FRK_ConfigScratch".Maximum, MaxLength := "FRK_ConfigScratch".MaxLength, Value := "FRK_ConfigScratch".Value);
           IF NOT #Ok THEN
               RETURN;
           END_IF;
           #Ok := "FRK_ConfigPut"(Scope := #Module.Status.Name, ModelCode := #Code, Text := #Request.TextValue, RootIndex := #RootIndex);
           IF NOT #Ok THEN
               RETURN;
           END_IF;
           IF NOT #Inactive THEN
               #Module.ParCfg.Timeout := DINT_TO_TIME(LINT_TO_DINT("FRK_ConfigScratch".Value.Number));
           END_IF;
           #FRK_CfgWrite_DeclarationCylinder := TRUE;
           RETURN;
       END_IF;
       "FRK_CfgDef_DeclarationCylinder"(FieldIndex := 2);
       IF #Request.NameValue = "FRK_ConfigScratch".Entry.WriteKey THEN
           #Matched := TRUE;
           IF DINT_TO_UDINT(#Request.IntValue) <> "FRK_ConfigScratch".Entry.WriteRevision THEN
               RETURN;
           END_IF;
           #Level := MAX(IN1 := #Access.Policy.Required[1], IN2 := "FRK_ConfigScratch".MinWrite);
           IF #Access.CurrentLevel < #Level THEN
               RETURN;
           END_IF;
           IF #Request.DurationMs <> 0 THEN
               RETURN;
           END_IF;
           #Code := "FRK_ConfigModelCode"(RootIndex := #RootIndex, ModelIndex := #Request.DurationMs);
           #Inactive := #Code <> "FRK_ConfigStore".ActiveModels[#RootIndex];
           IF "FRK_ConfigScratch".Entry.RequiresReady AND NOT #Inactive AND NOT #RootReady THEN
               RETURN;
           END_IF;
           #Ok := "FRK_ConfigDecode"(Text := #Request.TextValue, Storage := "FRK_ConfigScratch".Storage, Minimum := "FRK_ConfigScratch".Minimum, Maximum := "FRK_ConfigScratch".Maximum, MaxLength := "FRK_ConfigScratch".MaxLength, Value := "FRK_ConfigScratch".Value);
           IF NOT #Ok THEN
               RETURN;
           END_IF;
           #Ok := "FRK_ConfigPut"(Scope := #Module.Status.Name, ModelCode := #Code, Text := #Request.TextValue, RootIndex := #RootIndex);
           IF NOT #Ok THEN
               RETURN;
           END_IF;
           IF NOT #Inactive THEN
               #Module.ParCfg.Preset := LINT_TO_DINT("FRK_ConfigScratch".Value.Number);
           END_IF;
           #FRK_CfgWrite_DeclarationCylinder := TRUE;
           RETURN;
       END_IF;
   END_IF;
END_FUNCTION

FUNCTION "FRK_CfgWrite_DeclarationUnit" : Bool   // FC160, SCL
{ S7_Optimized_Access := 'TRUE' }
VERSION : 0.1
// stored: AutoNumber true, IsIECCheckEnabled false, SetENOAutomatically false, UDAEnableTagReadback false
   VAR_INPUT
      Request : "ST_HmiRequest";
      Access : "FRK_Access";
      RootIndex : Int;
      RootReady : Bool;
   END_VAR
   VAR_IN_OUT
      Core : "FRK_Core";
      Status : "ST_ModuleStatus";
      ParCfg : "ST_DeclarationParCfg";
      StationCfg : "ST_UnitProbeStationCfg";
      Cell : "FB_DeclarationCell";
      Satellite : "FB_SatelliteUnit";
      Matched : Bool;
   END_VAR
   VAR_TEMP
      Ok : Bool;
      Level : DInt;
      Code : String[64];
      Inactive : Bool;
   END_VAR
BEGIN

   #FRK_CfgWrite_DeclarationUnit := FALSE;
   IF #Request.TargetPath = STRING_TO_WSTRING(#Status.Name) OR (#Request.TargetPath = WSTRING#'' AND #Core.ParentIndex = 0) THEN
       "FRK_CfgDef_DeclarationUnit"(FieldIndex := 1);
       IF #Request.NameValue = "FRK_ConfigScratch".Entry.WriteKey THEN
           #Matched := TRUE;
           IF DINT_TO_UDINT(#Request.IntValue) <> "FRK_ConfigScratch".Entry.WriteRevision THEN
               RETURN;
           END_IF;
           #Level := MAX(IN1 := #Access.Policy.Required[1], IN2 := "FRK_ConfigScratch".MinWrite);
           IF #Access.CurrentLevel < #Level THEN
               RETURN;
           END_IF;
           IF #Request.DurationMs <> 0 AND #Core.ParentIndex <> 0 THEN
               RETURN;
           END_IF;
           #Code := "FRK_ConfigModelCode"(RootIndex := #RootIndex, ModelIndex := #Request.DurationMs);
           #Inactive := #Code <> "FRK_ConfigStore".ActiveModels[#RootIndex];
           IF "FRK_ConfigScratch".Entry.RequiresReady AND NOT #Inactive AND NOT #RootReady THEN
               RETURN;
           END_IF;
           #Ok := "FRK_ConfigDecode"(Text := #Request.TextValue, Storage := "FRK_ConfigScratch".Storage, Minimum := "FRK_ConfigScratch".Minimum, Maximum := "FRK_ConfigScratch".Maximum, MaxLength := "FRK_ConfigScratch".MaxLength, Value := "FRK_ConfigScratch".Value);
           IF NOT #Ok THEN
               RETURN;
           END_IF;
           #Ok := "FRK_ConfigPut"(Scope := #Status.Name, ModelCode := #Code, Text := #Request.TextValue, RootIndex := #RootIndex);
           IF NOT #Ok THEN
               RETURN;
           END_IF;
           IF NOT #Inactive THEN
               #ParCfg.Timeout := DINT_TO_TIME(LINT_TO_DINT("FRK_ConfigScratch".Value.Number));
           END_IF;
           #FRK_CfgWrite_DeclarationUnit := TRUE;
           RETURN;
       END_IF;
       "FRK_CfgDef_DeclarationUnit"(FieldIndex := 2);
       IF #Request.NameValue = "FRK_ConfigScratch".Entry.WriteKey THEN
           #Matched := TRUE;
           IF DINT_TO_UDINT(#Request.IntValue) <> "FRK_ConfigScratch".Entry.WriteRevision THEN
               RETURN;
           END_IF;
           #Level := MAX(IN1 := #Access.Policy.Required[1], IN2 := "FRK_ConfigScratch".MinWrite);
           IF #Access.CurrentLevel < #Level THEN
               RETURN;
           END_IF;
           IF #Request.DurationMs <> 0 AND #Core.ParentIndex <> 0 THEN
               RETURN;
           END_IF;
           #Code := "FRK_ConfigModelCode"(RootIndex := #RootIndex, ModelIndex := #Request.DurationMs);
           #Inactive := #Code <> "FRK_ConfigStore".ActiveModels[#RootIndex];
           IF "FRK_ConfigScratch".Entry.RequiresReady AND NOT #Inactive AND NOT #RootReady THEN
               RETURN;
           END_IF;
           #Ok := "FRK_ConfigDecode"(Text := #Request.TextValue, Storage := "FRK_ConfigScratch".Storage, Minimum := "FRK_ConfigScratch".Minimum, Maximum := "FRK_ConfigScratch".Maximum, MaxLength := "FRK_ConfigScratch".MaxLength, Value := "FRK_ConfigScratch".Value);
           IF NOT #Ok THEN
               RETURN;
           END_IF;
           #Ok := "FRK_ConfigPut"(Scope := #Status.Name, ModelCode := #Code, Text := #Request.TextValue, RootIndex := #RootIndex);
           IF NOT #Ok THEN
               RETURN;
           END_IF;
           IF NOT #Inactive THEN
               #ParCfg.Preset := LINT_TO_DINT("FRK_ConfigScratch".Value.Number);
           END_IF;
           #FRK_CfgWrite_DeclarationUnit := TRUE;
           RETURN;
       END_IF;
       "FRK_CfgDef_DeclarationUnit"(FieldIndex := 3);
       IF #Request.NameValue = "FRK_ConfigScratch".Entry.WriteKey THEN
           #Matched := TRUE;
           IF DINT_TO_UDINT(#Request.IntValue) <> "FRK_ConfigScratch".Entry.WriteRevision THEN
               RETURN;
           END_IF;
           #Level := MAX(IN1 := #Access.Policy.Required[1], IN2 := "FRK_ConfigScratch".MinWrite);
           IF #Access.CurrentLevel < #Level THEN
               RETURN;
           END_IF;
           IF #Request.DurationMs <> 0 THEN
               RETURN;
           END_IF;
           #Code := '';
           #Inactive := FALSE;
           IF "FRK_ConfigScratch".Entry.RequiresReady AND NOT #Inactive AND NOT #RootReady THEN
               RETURN;
           END_IF;
           #Ok := "FRK_ConfigDecode"(Text := #Request.TextValue, Storage := "FRK_ConfigScratch".Storage, Minimum := "FRK_ConfigScratch".Minimum, Maximum := "FRK_ConfigScratch".Maximum, MaxLength := "FRK_ConfigScratch".MaxLength, Value := "FRK_ConfigScratch".Value);
           IF NOT #Ok THEN
               RETURN;
           END_IF;
           #Ok := "FRK_ConfigPut"(Scope := #Status.Name, ModelCode := #Code, Text := #Request.TextValue, RootIndex := #RootIndex);
           IF NOT #Ok THEN
               RETURN;
           END_IF;
           IF NOT #Inactive THEN
               #StationCfg.SiteLabel := "FRK_ConfigScratch".Value.Text;
           END_IF;
           #FRK_CfgWrite_DeclarationUnit := TRUE;
           RETURN;
       END_IF;
       "FRK_CfgDef_DeclarationUnit"(FieldIndex := 4);
       IF #Request.NameValue = "FRK_ConfigScratch".Entry.WriteKey THEN
           #Matched := TRUE;
           IF DINT_TO_UDINT(#Request.IntValue) <> "FRK_ConfigScratch".Entry.WriteRevision THEN
               RETURN;
           END_IF;
           #Level := MAX(IN1 := #Access.Policy.Required[1], IN2 := "FRK_ConfigScratch".MinWrite);
           IF #Access.CurrentLevel < #Level THEN
               RETURN;
           END_IF;
           IF #Request.DurationMs <> 0 THEN
               RETURN;
           END_IF;
           #Code := '';
           #Inactive := FALSE;
           IF "FRK_ConfigScratch".Entry.RequiresReady AND NOT #Inactive AND NOT #RootReady THEN
               RETURN;
           END_IF;
           #Ok := "FRK_ConfigDecode"(Text := #Request.TextValue, Storage := "FRK_ConfigScratch".Storage, Minimum := "FRK_ConfigScratch".Minimum, Maximum := "FRK_ConfigScratch".Maximum, MaxLength := "FRK_ConfigScratch".MaxLength, Value := "FRK_ConfigScratch".Value);
           IF NOT #Ok THEN
               RETURN;
           END_IF;
           #Ok := "FRK_ConfigPut"(Scope := #Status.Name, ModelCode := #Code, Text := #Request.TextValue, RootIndex := #RootIndex);
           IF NOT #Ok THEN
               RETURN;
           END_IF;
           IF NOT #Inactive THEN
               #StationCfg.LongText := "FRK_ConfigScratch".Value.Text;
           END_IF;
           #FRK_CfgWrite_DeclarationUnit := TRUE;
           RETURN;
       END_IF;
       "FRK_CfgDef_DeclarationUnit"(FieldIndex := 5);
       IF #Request.NameValue = "FRK_ConfigScratch".Entry.WriteKey THEN
           #Matched := TRUE;
           IF DINT_TO_UDINT(#Request.IntValue) <> "FRK_ConfigScratch".Entry.WriteRevision THEN
               RETURN;
           END_IF;
           #Level := MAX(IN1 := #Access.Policy.Required[1], IN2 := "FRK_ConfigScratch".MinWrite);
           IF #Access.CurrentLevel < #Level THEN
               RETURN;
           END_IF;
           IF #Request.DurationMs <> 0 THEN
               RETURN;
           END_IF;
           #Code := '';
           #Inactive := FALSE;
           IF "FRK_ConfigScratch".Entry.RequiresReady AND NOT #Inactive AND NOT #RootReady THEN
               RETURN;
           END_IF;
           #Ok := "FRK_ConfigDecode"(Text := #Request.TextValue, Storage := "FRK_ConfigScratch".Storage, Minimum := "FRK_ConfigScratch".Minimum, Maximum := "FRK_ConfigScratch".Maximum, MaxLength := "FRK_ConfigScratch".MaxLength, Value := "FRK_ConfigScratch".Value);
           IF NOT #Ok THEN
               RETURN;
           END_IF;
           #Ok := "FRK_ConfigPut"(Scope := #Status.Name, ModelCode := #Code, Text := #Request.TextValue, RootIndex := #RootIndex);
           IF NOT #Ok THEN
               RETURN;
           END_IF;
           IF NOT #Inactive THEN
               #StationCfg.Enabled := "FRK_ConfigScratch".Value.Flag;
           END_IF;
           #FRK_CfgWrite_DeclarationUnit := TRUE;
           RETURN;
       END_IF;
   END_IF;
   #Ok := "FRK_CfgWrite_DeclarationCell"(Module := #Cell, Access := #Access, Request := #Request, RootIndex := #RootIndex, RootReady := #RootReady, Matched := #Matched);
   IF #Matched THEN
       #FRK_CfgWrite_DeclarationUnit := #Ok;
       RETURN;
   END_IF;
   #Ok := "FRK_CfgWrite_SatelliteUnit"(Module := #Satellite, Access := #Access, Request := #Request, RootIndex := #RootIndex, RootReady := #RootReady, Matched := #Matched);
   IF #Matched THEN
       #FRK_CfgWrite_DeclarationUnit := #Ok;
       RETURN;
   END_IF;
END_FUNCTION

FUNCTION "FRK_CfgWrite_InnerUnit" : Bool   // FC144, SCL
{ S7_Optimized_Access := 'TRUE' }
VERSION : 0.1
// stored: AutoNumber true, IsIECCheckEnabled false, SetENOAutomatically false, UDAEnableTagReadback false
   VAR_INPUT
      Request : "ST_HmiRequest";
      Access : "FRK_Access";
      RootIndex : Int;
      RootReady : Bool;
   END_VAR
   VAR_IN_OUT
      Module : "FB_InnerUnit";
      Matched : Bool;
   END_VAR
   VAR_TEMP
      Ok : Bool;
      Level : DInt;
      Code : String[64];
      Inactive : Bool;
   END_VAR
BEGIN

   #FRK_CfgWrite_InnerUnit := FALSE;
   IF #Request.TargetPath = STRING_TO_WSTRING(#Module.Status.Name) OR (#Request.TargetPath = WSTRING#'' AND #Module.Core.ParentIndex = 0) THEN
       "FRK_CfgDef_InnerUnit"(FieldIndex := 1);
       IF #Request.NameValue = "FRK_ConfigScratch".Entry.WriteKey THEN
           #Matched := TRUE;
           IF DINT_TO_UDINT(#Request.IntValue) <> "FRK_ConfigScratch".Entry.WriteRevision THEN
               RETURN;
           END_IF;
           #Level := MAX(IN1 := #Access.Policy.Required[1], IN2 := "FRK_ConfigScratch".MinWrite);
           IF #Access.CurrentLevel < #Level THEN
               RETURN;
           END_IF;
           IF #Request.DurationMs <> 0 THEN
               RETURN;
           END_IF;
           #Code := "FRK_ConfigModelCode"(RootIndex := #RootIndex, ModelIndex := #Request.DurationMs);
           #Inactive := #Code <> "FRK_ConfigStore".ActiveModels[#RootIndex];
           IF "FRK_ConfigScratch".Entry.RequiresReady AND NOT #Inactive AND NOT #RootReady THEN
               RETURN;
           END_IF;
           #Ok := "FRK_ConfigDecode"(Text := #Request.TextValue, Storage := "FRK_ConfigScratch".Storage, Minimum := "FRK_ConfigScratch".Minimum, Maximum := "FRK_ConfigScratch".Maximum, MaxLength := "FRK_ConfigScratch".MaxLength, Value := "FRK_ConfigScratch".Value);
           IF NOT #Ok THEN
               RETURN;
           END_IF;
           #Ok := "FRK_ConfigPut"(Scope := #Module.Status.Name, ModelCode := #Code, Text := #Request.TextValue, RootIndex := #RootIndex);
           IF NOT #Ok THEN
               RETURN;
           END_IF;
           IF NOT #Inactive THEN
               #Module.ParCfg.Timeout := DINT_TO_TIME(LINT_TO_DINT("FRK_ConfigScratch".Value.Number));
           END_IF;
           #FRK_CfgWrite_InnerUnit := TRUE;
           RETURN;
       END_IF;
       "FRK_CfgDef_InnerUnit"(FieldIndex := 2);
       IF #Request.NameValue = "FRK_ConfigScratch".Entry.WriteKey THEN
           #Matched := TRUE;
           IF DINT_TO_UDINT(#Request.IntValue) <> "FRK_ConfigScratch".Entry.WriteRevision THEN
               RETURN;
           END_IF;
           #Level := MAX(IN1 := #Access.Policy.Required[1], IN2 := "FRK_ConfigScratch".MinWrite);
           IF #Access.CurrentLevel < #Level THEN
               RETURN;
           END_IF;
           IF #Request.DurationMs <> 0 THEN
               RETURN;
           END_IF;
           #Code := "FRK_ConfigModelCode"(RootIndex := #RootIndex, ModelIndex := #Request.DurationMs);
           #Inactive := #Code <> "FRK_ConfigStore".ActiveModels[#RootIndex];
           IF "FRK_ConfigScratch".Entry.RequiresReady AND NOT #Inactive AND NOT #RootReady THEN
               RETURN;
           END_IF;
           #Ok := "FRK_ConfigDecode"(Text := #Request.TextValue, Storage := "FRK_ConfigScratch".Storage, Minimum := "FRK_ConfigScratch".Minimum, Maximum := "FRK_ConfigScratch".Maximum, MaxLength := "FRK_ConfigScratch".MaxLength, Value := "FRK_ConfigScratch".Value);
           IF NOT #Ok THEN
               RETURN;
           END_IF;
           #Ok := "FRK_ConfigPut"(Scope := #Module.Status.Name, ModelCode := #Code, Text := #Request.TextValue, RootIndex := #RootIndex);
           IF NOT #Ok THEN
               RETURN;
           END_IF;
           IF NOT #Inactive THEN
               #Module.ParCfg.Preset := LINT_TO_DINT("FRK_ConfigScratch".Value.Number);
           END_IF;
           #FRK_CfgWrite_InnerUnit := TRUE;
           RETURN;
       END_IF;
       "FRK_CfgDef_InnerUnit"(FieldIndex := 3);
       IF #Request.NameValue = "FRK_ConfigScratch".Entry.WriteKey THEN
           #Matched := TRUE;
           IF DINT_TO_UDINT(#Request.IntValue) <> "FRK_ConfigScratch".Entry.WriteRevision THEN
               RETURN;
           END_IF;
           #Level := MAX(IN1 := #Access.Policy.Required[1], IN2 := "FRK_ConfigScratch".MinWrite);
           IF #Access.CurrentLevel < #Level THEN
               RETURN;
           END_IF;
           IF #Request.DurationMs <> 0 THEN
               RETURN;
           END_IF;
           #Code := '';
           #Inactive := FALSE;
           IF "FRK_ConfigScratch".Entry.RequiresReady AND NOT #Inactive AND NOT #RootReady THEN
               RETURN;
           END_IF;
           #Ok := "FRK_ConfigDecode"(Text := #Request.TextValue, Storage := "FRK_ConfigScratch".Storage, Minimum := "FRK_ConfigScratch".Minimum, Maximum := "FRK_ConfigScratch".Maximum, MaxLength := "FRK_ConfigScratch".MaxLength, Value := "FRK_ConfigScratch".Value);
           IF NOT #Ok THEN
               RETURN;
           END_IF;
           #Ok := "FRK_ConfigPut"(Scope := #Module.Status.Name, ModelCode := #Code, Text := #Request.TextValue, RootIndex := #RootIndex);
           IF NOT #Ok THEN
               RETURN;
           END_IF;
           IF NOT #Inactive THEN
               #Module.StationCfg.SiteLabel := "FRK_ConfigScratch".Value.Text;
           END_IF;
           #FRK_CfgWrite_InnerUnit := TRUE;
           RETURN;
       END_IF;
       "FRK_CfgDef_InnerUnit"(FieldIndex := 4);
       IF #Request.NameValue = "FRK_ConfigScratch".Entry.WriteKey THEN
           #Matched := TRUE;
           IF DINT_TO_UDINT(#Request.IntValue) <> "FRK_ConfigScratch".Entry.WriteRevision THEN
               RETURN;
           END_IF;
           #Level := MAX(IN1 := #Access.Policy.Required[1], IN2 := "FRK_ConfigScratch".MinWrite);
           IF #Access.CurrentLevel < #Level THEN
               RETURN;
           END_IF;
           IF #Request.DurationMs <> 0 THEN
               RETURN;
           END_IF;
           #Code := '';
           #Inactive := FALSE;
           IF "FRK_ConfigScratch".Entry.RequiresReady AND NOT #Inactive AND NOT #RootReady THEN
               RETURN;
           END_IF;
           #Ok := "FRK_ConfigDecode"(Text := #Request.TextValue, Storage := "FRK_ConfigScratch".Storage, Minimum := "FRK_ConfigScratch".Minimum, Maximum := "FRK_ConfigScratch".Maximum, MaxLength := "FRK_ConfigScratch".MaxLength, Value := "FRK_ConfigScratch".Value);
           IF NOT #Ok THEN
               RETURN;
           END_IF;
           #Ok := "FRK_ConfigPut"(Scope := #Module.Status.Name, ModelCode := #Code, Text := #Request.TextValue, RootIndex := #RootIndex);
           IF NOT #Ok THEN
               RETURN;
           END_IF;
           IF NOT #Inactive THEN
               #Module.StationCfg.LongText := "FRK_ConfigScratch".Value.Text;
           END_IF;
           #FRK_CfgWrite_InnerUnit := TRUE;
           RETURN;
       END_IF;
       "FRK_CfgDef_InnerUnit"(FieldIndex := 5);
       IF #Request.NameValue = "FRK_ConfigScratch".Entry.WriteKey THEN
           #Matched := TRUE;
           IF DINT_TO_UDINT(#Request.IntValue) <> "FRK_ConfigScratch".Entry.WriteRevision THEN
               RETURN;
           END_IF;
           #Level := MAX(IN1 := #Access.Policy.Required[1], IN2 := "FRK_ConfigScratch".MinWrite);
           IF #Access.CurrentLevel < #Level THEN
               RETURN;
           END_IF;
           IF #Request.DurationMs <> 0 THEN
               RETURN;
           END_IF;
           #Code := '';
           #Inactive := FALSE;
           IF "FRK_ConfigScratch".Entry.RequiresReady AND NOT #Inactive AND NOT #RootReady THEN
               RETURN;
           END_IF;
           #Ok := "FRK_ConfigDecode"(Text := #Request.TextValue, Storage := "FRK_ConfigScratch".Storage, Minimum := "FRK_ConfigScratch".Minimum, Maximum := "FRK_ConfigScratch".Maximum, MaxLength := "FRK_ConfigScratch".MaxLength, Value := "FRK_ConfigScratch".Value);
           IF NOT #Ok THEN
               RETURN;
           END_IF;
           #Ok := "FRK_ConfigPut"(Scope := #Module.Status.Name, ModelCode := #Code, Text := #Request.TextValue, RootIndex := #RootIndex);
           IF NOT #Ok THEN
               RETURN;
           END_IF;
           IF NOT #Inactive THEN
               #Module.StationCfg.Enabled := "FRK_ConfigScratch".Value.Flag;
           END_IF;
           #FRK_CfgWrite_InnerUnit := TRUE;
           RETURN;
       END_IF;
   END_IF;
   #Ok := "FRK_CfgWrite_DeclarationCell"(Module := #Module.Cell, Access := #Access, Request := #Request, RootIndex := #RootIndex, RootReady := #RootReady, Matched := #Matched);
   IF #Matched THEN
       #FRK_CfgWrite_InnerUnit := #Ok;
       RETURN;
   END_IF;
END_FUNCTION

FUNCTION "FRK_CfgWrite_SatelliteUnit" : Bool   // FC152, SCL
{ S7_Optimized_Access := 'TRUE' }
VERSION : 0.1
// stored: AutoNumber true, IsIECCheckEnabled false, SetENOAutomatically false, UDAEnableTagReadback false
   VAR_INPUT
      Request : "ST_HmiRequest";
      Access : "FRK_Access";
      RootIndex : Int;
      RootReady : Bool;
   END_VAR
   VAR_IN_OUT
      Module : "FB_SatelliteUnit";
      Matched : Bool;
   END_VAR
   VAR_TEMP
      Ok : Bool;
      Level : DInt;
      Code : String[64];
      Inactive : Bool;
   END_VAR
BEGIN

   #FRK_CfgWrite_SatelliteUnit := FALSE;
   IF #Request.TargetPath = STRING_TO_WSTRING(#Module.Status.Name) OR (#Request.TargetPath = WSTRING#'' AND #Module.Core.ParentIndex = 0) THEN
       "FRK_CfgDef_SatelliteUnit"(FieldIndex := 1);
       IF #Request.NameValue = "FRK_ConfigScratch".Entry.WriteKey THEN
           #Matched := TRUE;
           IF DINT_TO_UDINT(#Request.IntValue) <> "FRK_ConfigScratch".Entry.WriteRevision THEN
               RETURN;
           END_IF;
           #Level := MAX(IN1 := #Access.Policy.Required[1], IN2 := "FRK_ConfigScratch".MinWrite);
           IF #Access.CurrentLevel < #Level THEN
               RETURN;
           END_IF;
           IF #Request.DurationMs <> 0 THEN
               RETURN;
           END_IF;
           #Code := "FRK_ConfigModelCode"(RootIndex := #RootIndex, ModelIndex := #Request.DurationMs);
           #Inactive := #Code <> "FRK_ConfigStore".ActiveModels[#RootIndex];
           IF "FRK_ConfigScratch".Entry.RequiresReady AND NOT #Inactive AND NOT #RootReady THEN
               RETURN;
           END_IF;
           #Ok := "FRK_ConfigDecode"(Text := #Request.TextValue, Storage := "FRK_ConfigScratch".Storage, Minimum := "FRK_ConfigScratch".Minimum, Maximum := "FRK_ConfigScratch".Maximum, MaxLength := "FRK_ConfigScratch".MaxLength, Value := "FRK_ConfigScratch".Value);
           IF NOT #Ok THEN
               RETURN;
           END_IF;
           #Ok := "FRK_ConfigPut"(Scope := #Module.Status.Name, ModelCode := #Code, Text := #Request.TextValue, RootIndex := #RootIndex);
           IF NOT #Ok THEN
               RETURN;
           END_IF;
           IF NOT #Inactive THEN
               #Module.ParCfg.Timeout := DINT_TO_TIME(LINT_TO_DINT("FRK_ConfigScratch".Value.Number));
           END_IF;
           #FRK_CfgWrite_SatelliteUnit := TRUE;
           RETURN;
       END_IF;
       "FRK_CfgDef_SatelliteUnit"(FieldIndex := 2);
       IF #Request.NameValue = "FRK_ConfigScratch".Entry.WriteKey THEN
           #Matched := TRUE;
           IF DINT_TO_UDINT(#Request.IntValue) <> "FRK_ConfigScratch".Entry.WriteRevision THEN
               RETURN;
           END_IF;
           #Level := MAX(IN1 := #Access.Policy.Required[1], IN2 := "FRK_ConfigScratch".MinWrite);
           IF #Access.CurrentLevel < #Level THEN
               RETURN;
           END_IF;
           IF #Request.DurationMs <> 0 THEN
               RETURN;
           END_IF;
           #Code := "FRK_ConfigModelCode"(RootIndex := #RootIndex, ModelIndex := #Request.DurationMs);
           #Inactive := #Code <> "FRK_ConfigStore".ActiveModels[#RootIndex];
           IF "FRK_ConfigScratch".Entry.RequiresReady AND NOT #Inactive AND NOT #RootReady THEN
               RETURN;
           END_IF;
           #Ok := "FRK_ConfigDecode"(Text := #Request.TextValue, Storage := "FRK_ConfigScratch".Storage, Minimum := "FRK_ConfigScratch".Minimum, Maximum := "FRK_ConfigScratch".Maximum, MaxLength := "FRK_ConfigScratch".MaxLength, Value := "FRK_ConfigScratch".Value);
           IF NOT #Ok THEN
               RETURN;
           END_IF;
           #Ok := "FRK_ConfigPut"(Scope := #Module.Status.Name, ModelCode := #Code, Text := #Request.TextValue, RootIndex := #RootIndex);
           IF NOT #Ok THEN
               RETURN;
           END_IF;
           IF NOT #Inactive THEN
               #Module.ParCfg.Preset := LINT_TO_DINT("FRK_ConfigScratch".Value.Number);
           END_IF;
           #FRK_CfgWrite_SatelliteUnit := TRUE;
           RETURN;
       END_IF;
       "FRK_CfgDef_SatelliteUnit"(FieldIndex := 3);
       IF #Request.NameValue = "FRK_ConfigScratch".Entry.WriteKey THEN
           #Matched := TRUE;
           IF DINT_TO_UDINT(#Request.IntValue) <> "FRK_ConfigScratch".Entry.WriteRevision THEN
               RETURN;
           END_IF;
           #Level := MAX(IN1 := #Access.Policy.Required[1], IN2 := "FRK_ConfigScratch".MinWrite);
           IF #Access.CurrentLevel < #Level THEN
               RETURN;
           END_IF;
           IF #Request.DurationMs <> 0 THEN
               RETURN;
           END_IF;
           #Code := '';
           #Inactive := FALSE;
           IF "FRK_ConfigScratch".Entry.RequiresReady AND NOT #Inactive AND NOT #RootReady THEN
               RETURN;
           END_IF;
           #Ok := "FRK_ConfigDecode"(Text := #Request.TextValue, Storage := "FRK_ConfigScratch".Storage, Minimum := "FRK_ConfigScratch".Minimum, Maximum := "FRK_ConfigScratch".Maximum, MaxLength := "FRK_ConfigScratch".MaxLength, Value := "FRK_ConfigScratch".Value);
           IF NOT #Ok THEN
               RETURN;
           END_IF;
           #Ok := "FRK_ConfigPut"(Scope := #Module.Status.Name, ModelCode := #Code, Text := #Request.TextValue, RootIndex := #RootIndex);
           IF NOT #Ok THEN
               RETURN;
           END_IF;
           IF NOT #Inactive THEN
               #Module.StationCfg.SiteLabel := "FRK_ConfigScratch".Value.Text;
           END_IF;
           #FRK_CfgWrite_SatelliteUnit := TRUE;
           RETURN;
       END_IF;
       "FRK_CfgDef_SatelliteUnit"(FieldIndex := 4);
       IF #Request.NameValue = "FRK_ConfigScratch".Entry.WriteKey THEN
           #Matched := TRUE;
           IF DINT_TO_UDINT(#Request.IntValue) <> "FRK_ConfigScratch".Entry.WriteRevision THEN
               RETURN;
           END_IF;
           #Level := MAX(IN1 := #Access.Policy.Required[1], IN2 := "FRK_ConfigScratch".MinWrite);
           IF #Access.CurrentLevel < #Level THEN
               RETURN;
           END_IF;
           IF #Request.DurationMs <> 0 THEN
               RETURN;
           END_IF;
           #Code := '';
           #Inactive := FALSE;
           IF "FRK_ConfigScratch".Entry.RequiresReady AND NOT #Inactive AND NOT #RootReady THEN
               RETURN;
           END_IF;
           #Ok := "FRK_ConfigDecode"(Text := #Request.TextValue, Storage := "FRK_ConfigScratch".Storage, Minimum := "FRK_ConfigScratch".Minimum, Maximum := "FRK_ConfigScratch".Maximum, MaxLength := "FRK_ConfigScratch".MaxLength, Value := "FRK_ConfigScratch".Value);
           IF NOT #Ok THEN
               RETURN;
           END_IF;
           #Ok := "FRK_ConfigPut"(Scope := #Module.Status.Name, ModelCode := #Code, Text := #Request.TextValue, RootIndex := #RootIndex);
           IF NOT #Ok THEN
               RETURN;
           END_IF;
           IF NOT #Inactive THEN
               #Module.StationCfg.LongText := "FRK_ConfigScratch".Value.Text;
           END_IF;
           #FRK_CfgWrite_SatelliteUnit := TRUE;
           RETURN;
       END_IF;
       "FRK_CfgDef_SatelliteUnit"(FieldIndex := 5);
       IF #Request.NameValue = "FRK_ConfigScratch".Entry.WriteKey THEN
           #Matched := TRUE;
           IF DINT_TO_UDINT(#Request.IntValue) <> "FRK_ConfigScratch".Entry.WriteRevision THEN
               RETURN;
           END_IF;
           #Level := MAX(IN1 := #Access.Policy.Required[1], IN2 := "FRK_ConfigScratch".MinWrite);
           IF #Access.CurrentLevel < #Level THEN
               RETURN;
           END_IF;
           IF #Request.DurationMs <> 0 THEN
               RETURN;
           END_IF;
           #Code := '';
           #Inactive := FALSE;
           IF "FRK_ConfigScratch".Entry.RequiresReady AND NOT #Inactive AND NOT #RootReady THEN
               RETURN;
           END_IF;
           #Ok := "FRK_ConfigDecode"(Text := #Request.TextValue, Storage := "FRK_ConfigScratch".Storage, Minimum := "FRK_ConfigScratch".Minimum, Maximum := "FRK_ConfigScratch".Maximum, MaxLength := "FRK_ConfigScratch".MaxLength, Value := "FRK_ConfigScratch".Value);
           IF NOT #Ok THEN
               RETURN;
           END_IF;
           #Ok := "FRK_ConfigPut"(Scope := #Module.Status.Name, ModelCode := #Code, Text := #Request.TextValue, RootIndex := #RootIndex);
           IF NOT #Ok THEN
               RETURN;
           END_IF;
           IF NOT #Inactive THEN
               #Module.StationCfg.Enabled := "FRK_ConfigScratch".Value.Flag;
           END_IF;
           #FRK_CfgWrite_SatelliteUnit := TRUE;
           RETURN;
       END_IF;
   END_IF;
   #Ok := "FRK_CfgWrite_DeclarationCell"(Module := #Module.Cell, Access := #Access, Request := #Request, RootIndex := #RootIndex, RootReady := #RootReady, Matched := #Matched);
   IF #Matched THEN
       #FRK_CfgWrite_SatelliteUnit := #Ok;
       RETURN;
   END_IF;
   #Ok := "FRK_CfgWrite_InnerUnit"(Module := #Module.Inner, Access := #Access, Request := #Request, RootIndex := #RootIndex, RootReady := #RootReady, Matched := #Matched);
   IF #Matched THEN
       #FRK_CfgWrite_SatelliteUnit := #Ok;
       RETURN;
   END_IF;
END_FUNCTION

FUNCTION "FRK_ClearDiag" : Void   // FC6, SCL
{ S7_Optimized_Access := 'TRUE' }
VERSION : 0.1
// stored: AutoNumber true, IsIECCheckEnabled false, SetENOAutomatically false, UDAEnableTagReadback false
   VAR_IN_OUT
      Status : "ST_ModuleStatus";
   END_VAR
BEGIN

   #Status.Diagnostic.ReasonCode := 0;
   #Status.Diagnostic.SourcePath := WSTRING#'';
   #Status.Diagnostic.Description := WSTRING#'';
   #Status.Diagnostic.IoTag := '';
   #Status.Diagnostic.IoAddress := '';
   #Status.Diagnostic.Severity := 0;
   #Status.Diagnostic.Category := 0;
   #Status.Diagnostic.Since := LDT#1970-01-01-00:00:00.000000000;
   #Status.Diagnostic.TimeSynchronized := FALSE;
END_FUNCTION

FUNCTION "FRK_ClockTick" : Void   // FC4, SCL
{ S7_Optimized_Access := 'TRUE' }
VERSION : 0.1
// Shared command kernel v0.1. Core 2.2 / 6.1 / 3.14 / 8.11.
//  Generated enum/rationalization values come from Core authorities.
// stored: AutoNumber true, IsIECCheckEnabled false, SetENOAutomatically false, UDAEnableTagReadback false
   VAR_TEMP
      DeltaS : LReal;
   END_VAR
BEGIN

   #DeltaS := RUNTIME("FRK_Clock".Mem);
   IF #DeltaS < 0.0 OR #DeltaS > 60.0 THEN
       #DeltaS := 0.0;
   END_IF;
   "FRK_Clock".AccMs := "FRK_Clock".AccMs + #DeltaS * 1000.0;
   IF "FRK_Clock".AccMs >= 4294967296.0 THEN
       "FRK_Clock".AccMs := "FRK_Clock".AccMs - 4294967296.0;
   END_IF;
   "FRK_Clock".NowMs := TRUNC_UDINT("FRK_Clock".AccMs);
END_FUNCTION

FUNCTION "FRK_Complete" : Void   // FC14, SCL
{ S7_Optimized_Access := 'TRUE' }
VERSION : 0.1
// stored: AutoNumber true, IsIECCheckEnabled false, SetENOAutomatically false, UDAEnableTagReadback false
   VAR_IN_OUT
      Core : "FRK_Core";
      Status : "ST_ModuleStatus";
   END_VAR
BEGIN

   IF #Core.Exec = 1 THEN
       #Core.Exec := 2;
       #Core.Step := 0;
       #Core.Dispatch := FALSE;
       "FRK_ClearDiag"(Status := #Status);
   END_IF;
END_FUNCTION

FUNCTION "FRK_ConfigAppend" : Void   // FC25, SCL
{ S7_Optimized_Access := 'TRUE' }
VERSION : 0.1
// stored: AutoNumber true, IsIECCheckEnabled false, SetENOAutomatically false, UDAEnableTagReadback false
   VAR_INPUT
      Scope : String;
      Item : String;
      ValueText : WString;
      ValueType : DInt;
      ReadLevel : DInt;
      Readable : Bool;
   END_VAR
   VAR_IN_OUT
      Cursor : "FRK_ConfigCursor";
      Page : "ST_ConfigPage";
   END_VAR
   VAR_TEMP
      Slot : DInt;
   END_VAR
BEGIN

   #Slot := #Cursor.Position - #Cursor.First;
   #Cursor.Position := #Cursor.Position + 1;
   IF #Slot < 0 OR #Slot >= 16 THEN
       RETURN;
   END_IF;
   #Slot := #Slot + 1;
   #Page.Entries[#Slot].Scope := STRING_TO_WSTRING(#Scope);
   #Page.Entries[#Slot].Item := STRING_TO_WSTRING(#Item);
   #Page.Entries[#Slot].ValueType := #ValueType;
   #Page.Entries[#Slot].ReadLevel := #ReadLevel;
   #Page.Entries[#Slot].Readable := #Readable;
   IF #Readable THEN
       #Page.Entries[#Slot].ValueText := #ValueText;
   END_IF;
   #Page.EntryCount := DINT_TO_INT(#Slot);
END_FUNCTION

FUNCTION "FRK_ConfigAppendEntry" : Void   // FC100, SCL
{ S7_Optimized_Access := 'TRUE' }
VERSION : 0.1
// stored: AutoNumber true, IsIECCheckEnabled false, SetENOAutomatically false, UDAEnableTagReadback false
   VAR_IN_OUT
      Cursor : "FRK_ConfigCursor";
      Page : "ST_ConfigPage";
   END_VAR
   VAR_TEMP
      Slot : DInt;
   END_VAR
BEGIN

   #Slot := #Cursor.Position - #Cursor.First;
   #Cursor.Position := #Cursor.Position + 1;
   IF #Slot < 0 OR #Slot >= 16 THEN
       RETURN;
   END_IF;
   #Slot := #Slot + 1;
   #Page.Entries[#Slot] := "FRK_ConfigScratch".Entry;
   #Page.EntryCount := DINT_TO_INT(#Slot);
END_FUNCTION

FUNCTION "FRK_ConfigBegin" : Void   // FC24, SCL
{ S7_Optimized_Access := 'TRUE' }
VERSION : 0.1
// stored: AutoNumber true, IsIECCheckEnabled false, SetENOAutomatically false, UDAEnableTagReadback false
   VAR_INPUT
      PageIndex : DInt;
      Revision : UDInt;
   END_VAR
   VAR_IN_OUT
      Cursor : "FRK_ConfigCursor";
      Page : "ST_ConfigPage";
   END_VAR
   VAR_TEMP
      Index : Int;
   END_VAR
BEGIN

   #Cursor.Position := 0;
   #Cursor.First := 0;
   #Page.Revision := #Revision;
   #Page.PageIndex := 0;
   IF #PageIndex >= 0 AND #PageIndex <= 32767 THEN
       #Cursor.First := #PageIndex * 16;
       #Page.PageIndex := DINT_TO_INT(#PageIndex);
   END_IF;
   #Page.PageCount := 1;
   #Page.EntryCount := 0;
   "FRK_UnitScratch".EmptyConfigEntry.ValueType := 1;
   "FRK_UnitScratch".EmptyConfigEntry.Readable := TRUE;
   FOR #Index := 1 TO 16 DO
       #Page.Entries[#Index] := "FRK_UnitScratch".EmptyConfigEntry;
   END_FOR;
END_FUNCTION

FUNCTION "FRK_ConfigBoot" : Void   // FC104, SCL
{ S7_Optimized_Access := 'TRUE' }
VERSION : 0.1
// stored: AutoNumber true, IsIECCheckEnabled false, SetENOAutomatically false, UDAEnableTagReadback false
   VAR_INPUT
      Startup : Bool;
   END_VAR
   VAR_TEMP
      Index : Int;
   END_VAR
BEGIN

   IF NOT #Startup THEN
       RETURN;
   END_IF;
   "FRK_ConfigRuntime".Fresh := "FRK_ConfigStore".SchemaVersion = 0;
   IF "FRK_ConfigStore".SchemaVersion <> 1 THEN
       FOR #Index := 1 TO 114 DO
           "FRK_ConfigStore".Rows[#Index].Used := FALSE;
       END_FOR;
       IF NOT "FRK_ConfigRuntime".Fresh THEN
           "FRK_ConfigLoss"(RootIndex := 1,
                            Scope := 'StationA');
       END_IF;
       "FRK_ConfigStore".ActiveModels[1] := 'MODEL_A';
       IF NOT "FRK_ConfigRuntime".Fresh THEN
           "FRK_ConfigLoss"(RootIndex := 2,
                            Scope := 'StationB');
       END_IF;
       "FRK_ConfigStore".ActiveModels[2] := 'MODEL_A';
       "FRK_ConfigStore".SchemaVersion := 1;
   END_IF;
   IF "FRK_ConfigStore".ActiveModels[1] <> 'MODEL_A' AND "FRK_ConfigStore".ActiveModels[1] <> 'MODEL_B' THEN
       "FRK_ConfigStore".ActiveModels[1] := 'MODEL_A';
       "FRK_ConfigLoss"(RootIndex := 1,
                        Scope := 'StationA');
   END_IF;
   IF "FRK_ConfigStore".ActiveModels[2] <> 'MODEL_A' AND "FRK_ConfigStore".ActiveModels[2] <> 'MODEL_B' THEN
       "FRK_ConfigStore".ActiveModels[2] := 'MODEL_A';
       "FRK_ConfigLoss"(RootIndex := 2,
                        Scope := 'StationB');
   END_IF;
END_FUNCTION

FUNCTION "FRK_ConfigCatalog" : Void   // FC27, SCL
{ S7_Optimized_Access := 'TRUE' }
VERSION : 0.1
// stored: AutoNumber true, IsIECCheckEnabled false, SetENOAutomatically false, UDAEnableTagReadback false
   VAR_INPUT
      Scope : String;
      Count : Int;
      Catalog : Array[1..12] of "ST_CommandInfo";
      ReadLevel : DInt;
      Readable : Bool;
   END_VAR
   VAR_IN_OUT
      Cursor : "FRK_ConfigCursor";
      Page : "ST_ConfigPage";
   END_VAR
   VAR_TEMP
      Index : Int;
      IndexText : String[8];
      Prefix : String[254];
      Item : String[254];
   END_VAR
BEGIN

   "FRK_ConfigAppend"(Scope := #Scope,
                      Item := 'CatalogCount',
                      ValueText := STRING_TO_WSTRING(INT_TO_STRING(#Count)),
                      ValueType := 0,
                      ReadLevel := #ReadLevel,
                      Readable := #Readable,
                      Cursor := #Cursor,
                      Page := #Page);
   FOR #Index := 1 TO #Count DO
       IF #Index > 12 THEN
           EXIT;
       END_IF;
       #IndexText := INT_TO_STRING(#Index);
       IF #IndexText[1] = '+' THEN
           #IndexText := DELETE(IN := #IndexText, L := 1, P := 1);
       END_IF;
       #Prefix := CONCAT(IN1 := 'Catalog/Catalog[', IN2 := #IndexText);
       #Prefix := CONCAT(IN1 := #Prefix, IN2 := ']/');
       #Item := CONCAT(IN1 := #Prefix, IN2 := 'Value');
       "FRK_ConfigAppend"(Scope := #Scope,
                          Item := #Item,
                          ValueText := STRING_TO_WSTRING(DINT_TO_STRING(#Catalog[#Index].Value)),
                          ValueType := 0,
                          ReadLevel := #ReadLevel,
                          Readable := #Readable,
                          Cursor := #Cursor,
                          Page := #Page);
       #Item := CONCAT(IN1 := #Prefix, IN2 := 'Label');
       "FRK_ConfigAppend"(Scope := #Scope,
                          Item := #Item,
                          ValueText := STRING_TO_WSTRING(#Catalog[#Index].Label),
                          ValueType := 1,
                          ReadLevel := #ReadLevel,
                          Readable := #Readable,
                          Cursor := #Cursor,
                          Page := #Page);
       #Item := CONCAT(IN1 := #Prefix, IN2 := 'Style');
       "FRK_ConfigAppend"(Scope := #Scope,
                          Item := #Item,
                          ValueText := STRING_TO_WSTRING(DINT_TO_STRING(#Catalog[#Index].Style)),
                          ValueType := 0,
                          ReadLevel := #ReadLevel,
                          Readable := #Readable,
                          Cursor := #Cursor,
                          Page := #Page);
   END_FOR;
END_FUNCTION

FUNCTION "FRK_ConfigDecode" : Bool   // FC95, SCL
{ S7_Optimized_Access := 'TRUE' }
VERSION : 0.1
// Keyed local-retain config. The typed owner validates before publishing a value.
// stored: AutoNumber true, IsIECCheckEnabled false, SetENOAutomatically false, UDAEnableTagReadback false
   VAR_INPUT
      Text : WString;
      Storage : DInt;
      Minimum : LReal;
      Maximum : LReal;
      MaxLength : Int;
   END_VAR
   VAR_IN_OUT
      Value : "FRK_ConfigValue";
   END_VAR
   VAR_TEMP
      Index : Int;
      Width : Int;
      Negative : Bool;
      Magnitude : ULInt;
      Digit : ULInt;
   END_VAR
BEGIN

   #FRK_ConfigDecode := FALSE;
   IF #Storage = 8 THEN
       IF LEN(#Text) > #MaxLength THEN
           RETURN;
       END_IF;
       #Value.Text := WSTRING_TO_STRING(#Text);
       IF STRING_TO_WSTRING(#Value.Text) <> #Text THEN
           RETURN;
       END_IF;
       #FRK_ConfigDecode := TRUE;
       RETURN;
   END_IF;
   IF #Storage = 1 THEN
       IF #Text = WSTRING#'true' OR #Text = WSTRING#'TRUE' OR #Text = WSTRING#'1' THEN
           #Value.Flag := TRUE;
       ELSIF #Text = WSTRING#'false' OR #Text = WSTRING#'FALSE' OR #Text = WSTRING#'0' THEN
           #Value.Flag := FALSE;
       ELSE
           RETURN;
       END_IF;
       #FRK_ConfigDecode := TRUE;
       RETURN;
   END_IF;
   #Width := LEN(#Text);
   IF #Width = 0 THEN
       RETURN;
   END_IF;
   #Negative := FALSE;
   #Index := 1;
   IF #Text[1] = WCHAR#'-' THEN
       #Negative := TRUE;
       #Index := 2;
   ELSIF #Text[1] = WCHAR#'+' THEN
       #Index := 2;
   END_IF;
   IF #Index > #Width THEN
       RETURN;
   END_IF;
   #Magnitude := 0;
   WHILE #Index <= #Width DO
       IF #Text[#Index] < WCHAR#'0' OR #Text[#Index] > WCHAR#'9' THEN
           RETURN;
       END_IF;
       #Digit := UINT_TO_ULINT(WCHAR_TO_UINT(#Text[#Index]) - UINT#48);
       IF #Magnitude > (ULINT#4294967295 - #Digit) / ULINT#10 THEN
           RETURN;
       END_IF;
       #Magnitude := #Magnitude * ULINT#10 + #Digit;
       #Index := #Index + 1;
   END_WHILE;
   #Value.Number := ULINT_TO_LINT(#Magnitude);
   IF #Negative THEN
       #Value.Number := - #Value.Number;
   END_IF;
   IF LINT_TO_LREAL(#Value.Number) < #Minimum OR LINT_TO_LREAL(#Value.Number) > #Maximum THEN
       RETURN;
   END_IF;
   #FRK_ConfigDecode := TRUE;
END_FUNCTION

FUNCTION "FRK_ConfigFind" : Int   // FC96, SCL
{ S7_Optimized_Access := 'TRUE' }
VERSION : 0.1
// stored: AutoNumber true, IsIECCheckEnabled false, SetENOAutomatically false, UDAEnableTagReadback false
   VAR_INPUT
      Scope : String;
      Key : String;
      ModelCode : String;
   END_VAR
   VAR_TEMP
      Index : Int;
   END_VAR
BEGIN

   #FRK_ConfigFind := 0;
   FOR #Index := 1 TO 114 DO
       IF "FRK_ConfigStore".Rows[#Index].Used
           AND "FRK_ConfigStore".Rows[#Index].Record.Scope = #Scope
           AND "FRK_ConfigStore".Rows[#Index].Record.WriteKey = #Key
           AND "FRK_ConfigStore".Rows[#Index].ModelCode = #ModelCode THEN
           #FRK_ConfigFind := #Index;
           RETURN;
       END_IF;
   END_FOR;
END_FUNCTION

FUNCTION "FRK_ConfigFinish" : Void   // FC26, SCL
{ S7_Optimized_Access := 'TRUE' }
VERSION : 0.1
// stored: AutoNumber true, IsIECCheckEnabled false, SetENOAutomatically false, UDAEnableTagReadback false
   VAR_IN_OUT
      Cursor : "FRK_ConfigCursor";
      Page : "ST_ConfigPage";
   END_VAR
BEGIN

   #Page.PageCount := DINT_TO_INT((#Cursor.Position + 16 - 1) / 16);
   IF #Page.PageCount < 1 THEN
       #Page.PageCount := 1;
   END_IF;
END_FUNCTION

FUNCTION "FRK_ConfigGet" : Bool   // FC98, SCL
{ S7_Optimized_Access := 'TRUE' }
VERSION : 0.1
// stored: AutoNumber true, IsIECCheckEnabled false, SetENOAutomatically false, UDAEnableTagReadback false
   VAR_INPUT
      Scope : String;
      ModelCode : String;
   END_VAR
   VAR_TEMP
      Index : Int;
   END_VAR
BEGIN

   #FRK_ConfigGet := FALSE;
   #Index := "FRK_ConfigFind"(Scope := #Scope, Key := "FRK_ConfigScratch".Entry.WriteKey, ModelCode := #ModelCode);
   IF #Index = 0 THEN
       RETURN;
   END_IF;
   IF "FRK_ConfigStore".Rows[#Index].SchemaVersion <> "FRK_ConfigScratch".Schema
       OR "FRK_ConfigStore".Rows[#Index].Record.Revision <> "FRK_ConfigScratch".Entry.WriteRevision
       OR "FRK_ConfigStore".Rows[#Index].Record.Kind <> "FRK_ConfigScratch".Entry.ConfigKind
       OR "FRK_ConfigStore".Rows[#Index].Record.ValueType <> "FRK_ConfigScratch".Entry.ValueType THEN
       RETURN;
   END_IF;
   #FRK_ConfigGet := "FRK_ConfigDecode"(Text := STRING_TO_WSTRING("FRK_ConfigStore".Rows[#Index].Record.ValueText),
                                        Storage := "FRK_ConfigScratch".Storage, Minimum := "FRK_ConfigScratch".Minimum, Maximum := "FRK_ConfigScratch".Maximum,
                                        MaxLength := "FRK_ConfigScratch".MaxLength, Value := "FRK_ConfigScratch".Value);
   "FRK_ConfigScratch".Entry.ValueText := STRING_TO_WSTRING("FRK_ConfigStore".Rows[#Index].Record.ValueText);
END_FUNCTION

FUNCTION "FRK_ConfigLoss" : Void   // FC99, SCL
{ S7_Optimized_Access := 'TRUE' }
VERSION : 0.1
// stored: AutoNumber true, IsIECCheckEnabled false, SetENOAutomatically false, UDAEnableTagReadback false
   VAR_INPUT
      RootIndex : Int;
      Scope : String;
   END_VAR
BEGIN

   IF #RootIndex < 1 OR #RootIndex > 2 THEN
       RETURN;
   END_IF;
   "FRK_ConfigStore".Lost[#RootIndex] := TRUE;
   "FRK_ConfigStore".Acknowledged[#RootIndex] := FALSE;
   "FRK_ConfigStore".LostPath[#RootIndex] := #Scope;
END_FUNCTION

FUNCTION "FRK_ConfigModelCode" : String   // FC103, SCL
{ S7_Optimized_Access := 'TRUE' }
VERSION : 0.1
// stored: AutoNumber true, IsIECCheckEnabled false, SetENOAutomatically false, UDAEnableTagReadback false
   VAR_INPUT
      RootIndex : Int;
      ModelIndex : UDInt;
   END_VAR
BEGIN

   #FRK_ConfigModelCode := '';
   IF #RootIndex < 1 OR #RootIndex > 2 THEN
       RETURN;
   END_IF;
   IF #ModelIndex = 0 THEN
       #FRK_ConfigModelCode := "FRK_ConfigStore".ActiveModels[#RootIndex];
       RETURN;
   END_IF;
   CASE #ModelIndex OF
       1:
           #FRK_ConfigModelCode := 'MODEL_A';
       2:
           #FRK_ConfigModelCode := 'MODEL_B';
       ELSE
           RETURN;
   END_CASE;
END_FUNCTION

FUNCTION "FRK_ConfigPut" : Bool   // FC97, SCL
{ S7_Optimized_Access := 'TRUE' }
VERSION : 0.1
// stored: AutoNumber true, IsIECCheckEnabled false, SetENOAutomatically false, UDAEnableTagReadback false
   VAR_INPUT
      Scope : String;
      ModelCode : String;
      Text : WString;
      RootIndex : Int;
   END_VAR
   VAR_TEMP
      Index : Int;
   END_VAR
BEGIN

   #FRK_ConfigPut := FALSE;
   IF #RootIndex < 1 OR #RootIndex > 2 THEN
       RETURN;
   END_IF;
   IF "FRK_ConfigRuntime".Unavailable THEN
       "FRK_ConfigRuntime".Failed[#RootIndex] := TRUE;
       RETURN;
   END_IF;
   IF LEN(#Scope) > 80 OR LEN(#Text) > 80 THEN
       RETURN;
   END_IF;
   #Index := "FRK_ConfigFind"(Scope := #Scope, Key := "FRK_ConfigScratch".Entry.WriteKey, ModelCode := #ModelCode);
   IF #Index = 0 THEN
       FOR #Index := 1 TO 114 DO
           IF NOT "FRK_ConfigStore".Rows[#Index].Used THEN
               EXIT;
           END_IF;
       END_FOR;
   END_IF;
   IF #Index < 1 OR #Index > 114 THEN
       "FRK_ConfigRuntime".Failed[#RootIndex] := TRUE;
       RETURN;
   END_IF;
   "FRK_ConfigStore".Rows[#Index].SchemaVersion := "FRK_ConfigScratch".Schema;
   "FRK_ConfigStore".Rows[#Index].ModelCode := #ModelCode;
   "FRK_ConfigStore".Rows[#Index].Record.Scope := #Scope;
   "FRK_ConfigStore".Rows[#Index].Record.WriteKey := "FRK_ConfigScratch".Entry.WriteKey;
   "FRK_ConfigStore".Rows[#Index].Record.Revision := "FRK_ConfigScratch".Entry.WriteRevision;
   "FRK_ConfigStore".Rows[#Index].Record.Kind := "FRK_ConfigScratch".Entry.ConfigKind;
   "FRK_ConfigStore".Rows[#Index].Record.ValueType := "FRK_ConfigScratch".Entry.ValueType;
   "FRK_ConfigStore".Rows[#Index].Record.ValueText := WSTRING_TO_STRING(#Text);
   "FRK_ConfigStore".Rows[#Index].Used := TRUE;
   "FRK_ConfigRuntime".Failed[#RootIndex] := FALSE;
   #FRK_ConfigPut := TRUE;
END_FUNCTION

FUNCTION "FRK_ConfigRevision" : UDInt   // FC23, SCL
{ S7_Optimized_Access := 'TRUE' }
VERSION : 0.1
// Core 3.10.2: deterministic typed walk, one bounded response window.
//  Static facets carry no write capability. Every reused slot is cleared.
// stored: AutoNumber true, IsIECCheckEnabled false, SetENOAutomatically false, UDAEnableTagReadback false
   VAR_INPUT
      Previous : UDInt;
   END_VAR
   VAR_TEMP
      Stamp : DTL;
      ResultCode : Int;
      Generation : ULInt;
   END_VAR
BEGIN

   #FRK_ConfigRevision := #Previous + 1;
   #ResultCode := RD_SYS_T(OUT => #Stamp);
   IF #ResultCode = 0 THEN
       #Generation := LDT_TO_ULINT(DTL_TO_LDT(#Stamp)) / ULINT#1000000;
       #FRK_ConfigRevision := ULINT_TO_UDINT(#Generation MOD ULINT#4294967296);
   END_IF;
   IF #FRK_ConfigRevision = #Previous THEN
       #FRK_ConfigRevision := #Previous + 1;
   END_IF;
   IF #FRK_ConfigRevision = 0 THEN
       #FRK_ConfigRevision := 1;
   END_IF;
END_FUNCTION

FUNCTION "FRK_ConfigRoot" : Int   // FC102, SCL
{ S7_Optimized_Access := 'TRUE' }
VERSION : 0.1
// stored: AutoNumber true, IsIECCheckEnabled false, SetENOAutomatically false, UDAEnableTagReadback false
   VAR_INPUT
      RegIndex : DInt;
   END_VAR
BEGIN

   #FRK_ConfigRoot := 0;
   CASE #RegIndex OF
       1:
           #FRK_ConfigRoot := 1;
       2:
           #FRK_ConfigRoot := 1;
       3:
           #FRK_ConfigRoot := 1;
       4:
           #FRK_ConfigRoot := 1;
       5:
           #FRK_ConfigRoot := 1;
       6:
           #FRK_ConfigRoot := 1;
       7:
           #FRK_ConfigRoot := 1;
       8:
           #FRK_ConfigRoot := 1;
       9:
           #FRK_ConfigRoot := 1;
       10:
           #FRK_ConfigRoot := 1;
       11:
           #FRK_ConfigRoot := 1;
       12:
           #FRK_ConfigRoot := 1;
       13:
           #FRK_ConfigRoot := 2;
       14:
           #FRK_ConfigRoot := 2;
       15:
           #FRK_ConfigRoot := 2;
       16:
           #FRK_ConfigRoot := 2;
       17:
           #FRK_ConfigRoot := 2;
       18:
           #FRK_ConfigRoot := 2;
       19:
           #FRK_ConfigRoot := 2;
       20:
           #FRK_ConfigRoot := 2;
       21:
           #FRK_ConfigRoot := 2;
       22:
           #FRK_ConfigRoot := 2;
       23:
           #FRK_ConfigRoot := 2;
       24:
           #FRK_ConfigRoot := 2;
       ELSE
           RETURN;
   END_CASE;
END_FUNCTION

FUNCTION "FRK_ConfigStatus" : Void   // FC101, SCL
{ S7_Optimized_Access := 'TRUE' }
VERSION : 0.1
// stored: AutoNumber true, IsIECCheckEnabled false, SetENOAutomatically false, UDAEnableTagReadback false
   VAR_INPUT
      RootIndex : Int;
      Scope : String;
      PolicyLost : Bool;
      UsersLost : Bool;
   END_VAR
   VAR_IN_OUT
      Persist : "ST_ConfigPersistStatus";
      AlarmLog : "FRK_AlarmLog";
   END_VAR
   VAR_TEMP
      Diag : "ST_Diagnostic";
      Accepted : Bool;
   END_VAR
BEGIN

   IF #RootIndex < 1 OR #RootIndex > 2 THEN
       RETURN;
   END_IF;
   #Persist.Pending := FALSE;
   #Persist.Failed := "FRK_ConfigRuntime".Failed[#RootIndex];
   #Persist.StoreKind := 0;
   // Named set operations are not wired by the live retained-value provider.
   #Persist.StorePresent := TRUE;
   #Persist.RestoreLost := "FRK_ConfigStore".Lost[#RootIndex] OR #PolicyLost OR #UsersLost;
   #Persist.RestoreAcknowledged := "FRK_ConfigStore".Acknowledged[#RootIndex] AND NOT #PolicyLost AND NOT #UsersLost;
   IF #PolicyLost THEN
       #Persist.LostPath := CONCAT(IN1 := #Scope, IN2 := '.AccessPolicy');
   ELSIF #UsersLost THEN
       #Persist.LostPath := CONCAT(IN1 := #Scope, IN2 := '.Access');
   ELSE
       #Persist.LostPath := "FRK_ConfigStore".LostPath[#RootIndex];
   END_IF;
   // Access owns its precise loss events; announce only typed-config loss here.
   IF "FRK_ConfigStore".Lost[#RootIndex] AND NOT "FRK_ConfigStore".Acknowledged[#RootIndex] THEN
       IF "FRK_ConfigRuntime".LossSlot[#RootIndex] = 0 THEN
           #Diag := "FRK_UnitScratch".EmptyDiagnostic;
           #Diag.ReasonCode := 2040;
           #Diag.Description := WSTRING#'std.error.configRestoreLost';
           #Diag.SourcePath := STRING_TO_WSTRING("FRK_ConfigStore".LostPath[#RootIndex]);
           "FRK_ConfigRuntime".LossSlot[#RootIndex] := "FRK_AlarmRaise"(AlarmLog := #AlarmLog, Diag := #Diag, ResetClass := 0);
       END_IF;
   ELSIF "FRK_ConfigRuntime".LossSlot[#RootIndex] > 0 THEN
       #Accepted := "FRK_AlarmGone"(AlarmLog := #AlarmLog, Slot := "FRK_ConfigRuntime".LossSlot[#RootIndex]);
       "FRK_ConfigRuntime".LossSlot[#RootIndex] := 0;
   END_IF;
END_FUNCTION

FUNCTION "FRK_ConfigUnit" : Void   // FC28, SCL
{ S7_Optimized_Access := 'TRUE' }
VERSION : 0.1
// stored: AutoNumber true, IsIECCheckEnabled false, SetENOAutomatically false, UDAEnableTagReadback false
   VAR_INPUT
      Scope : String;
      Policy : Array[0..6] of "ST_ModePolicy";
      ModelCount : Int;
      ReadLevel : DInt;
      Readable : Bool;
   END_VAR
   VAR_IN_OUT
      Cursor : "FRK_ConfigCursor";
      Page : "ST_ConfigPage";
   END_VAR
   VAR_TEMP
      Index : Int;
      IndexText : String[8];
      Prefix : String[254];
      Item : String[254];
   END_VAR
BEGIN

